(* IEC 61131-3 sources: daoli-st-library/DL_MathData (part 24) *)

(* ---- FC_DL_StatsDevSumSq.st ---- *)
(*
  ============================================================
  组件名 : FC_DL_StatsDevSumSq
  分类   : DL_MathData
  功能   : 定长样本的离差平方和、自由度与方差计算，支持外部给定均值
  开源溯源 : internal-design（本轮无外部代码逐行引用）
             参考语义 : 无外部参考
  复杂度 : C1
  版本   : 1.0.0
  ============================================================
*)

FUNCTION FC_DL_StatsDevSumSq : REAL
VAR_INPUT
    aData        : ARRAY[0..31] OF REAL; // 样本数组，定长三十二 [工程单位] sample array of thirty two fixed slots [engineering unit]
    nCount       : INT; // 有效样本数 1~32 [个] effective sample count from one to thirty two [count]
    rMeanGiven   : REAL; // 外部给定的均值 [工程单位] externally supplied mean [engineering unit]
    bUseGivenMean: BOOL; // 真为使用给定均值，假为按样本自算 use the supplied mean when true
END_VAR
VAR_OUTPUT
    rSs    : REAL; // 离差平方和 [工程单位平方] sum of squared deviations [engineering unit squared]
    rDf    : REAL; // 自由度 [个] degrees of freedom [count]
    rVar   : REAL; // 方差 [工程单位平方] variance [engineering unit squared]
    bValid : BOOL; // 结果有效标志 result validity flag
END_VAR
VAR CONSTANT
    DL_CAP : INT := 32; // 数组容量 [个] array capacity [count]
END_VAR
VAR
    i      : INT := 0; // 遍历游标 [个] walk cursor [count]
    _rMean : REAL := 0.0; // 实际使用的均值 [工程单位] mean actually used [engineering unit]
    _rSum  : REAL := 0.0; // 样本和 [工程单位] sum of the samples [engineering unit]
    _rSs   : REAL := 0.0; // 平方和中间量 [工程单位平方] intermediate sum of squares [engineering unit squared]
    _rDev  : REAL := 0.0; // 单点离差 [工程单位] single deviation [engineering unit]
END_VAR

// 段 1｜出口预置 preset the exit
FC_DL_StatsDevSumSq := 0.0; // 缺省返回零 default zero return
rSs := 0.0; // 平方和预置零 sum of squares preset to zero
rDf := 0.0; // 自由度预置零 freedom preset to zero
rVar := 0.0; // 方差预置零 variance preset to zero
bValid := FALSE; // 计算完成前不认结果 unusable before the calculation
// 段 2｜点数闸与有限闸 count gate and finiteness gate
IF (nCount < 1) OR (nCount > DL_CAP) THEN
    RETURN; // 点数越界即无效 an out of range count is void
END_IF
IF (rMeanGiven <> rMeanGiven) OR ((aData[0] <> aData[0])) THEN
    RETURN; // 均值或首样本非有限即无效 a non finite mean or first sample is void
END_IF
// 段 3｜均值来源选择 the mean source selection
IF bUseGivenMean THEN
    _rMean := rMeanGiven; // 使用外部给定均值 use the supplied mean
ELSE
    _rSum := 0.0; // 样本和清零 clear the sum
    FOR i := 0 TO (nCount - 1) DO
        IF aData[i] <> aData[i] THEN
            RETURN; // 非有限样本拒收 refuse a non finite sample
        END_IF
        _rSum := _rSum + aData[i]; // 样本累加 accumulate the sample
    END_FOR
    _rMean := _rSum / INT_TO_REAL(nCount); // 自算均值，除子为已证正计数 the computed mean over a proven positive count
END_IF
// 段 4｜离差平方和 sum of squared deviations
_rSs := 0.0; // 平方和清零 clear the sum of squares
FOR i := 0 TO (nCount - 1) DO
    IF aData[i] <> aData[i] THEN
        RETURN; // 非有限样本拒收 refuse a non finite sample
    END_IF
    _rDev := aData[i] - _rMean; // 单点离差 single deviation
    _rSs := _rSs + _rDev * _rDev; // 平方累加 accumulate the square
END_FOR
rSs := _rSs; // 平方和落定 land the sum of squares
// 段 5｜自由度与方差自由度闸 freedom and the variance gate
rDf := INT_TO_REAL(nCount - 1); // 自由度取样本数减一 the freedom is the count minus one
IF rDf <= 0.0 THEN
    RETURN; // 自由度非正时方差不可求 a non positive freedom carries no variance
END_IF
rVar := _rSs / rDf; // 方差，除子为已证正自由度 variance over a proven positive freedom
bValid := TRUE; // 结果可用 result usable
FC_DL_StatsDevSumSq := _rSs; // 函数返回离差平方和 return the sum of squares
END_FUNCTION

(* ---- FC_DL_StatsEntropyCalc.st ---- *)
(*==============================================================================
 * 组件名称 : FC_DL_StatsEntropyCalc ｜ 子库 : DL_MathData ｜ v1.0.0 ｜ 2026-11-24
 * 平台     : CODESYS 3.5 / TwinCAT 3 / InoProShop / Machine Expert（纯 IEC，无厂商库）
 * 功能简介 : 香农熵 H = −Σ p·log2(p) [bit]，供直方图分布集中度、缺陷类别混杂度、
 *            多路料仓配比均匀度评估。概率先求和再归一化（q = p / Σp），故入参不要求
 *            严格和为 1（计数直方图可直接喂入）。
 * 契约     : 1 ≤ nCnt ≤ 8、各 p ≥ 0 且有限、Σp > 1.0E-12 → 返回 H ≥ 0、bValid := TRUE；
 *            nCnt 越界、任一 p 为负或非有限、Σp ≤ 1.0E-12（全零/近零，熵无定义）→
 *            返回 0、bError := TRUE、bValid := FALSE。
 * 依赖     : 无 DL_ 内部依赖（R16 自足实现），仅用标准库 LN；log2(p) 以 LN(p)/LN(2) 实现
 * 错误码   : R297 零码位范式：eErr 恒 0，仅以 bError / bValid 表达
 * 红线自检 : R1 零全局 R2 零%I/%Q R3 纯IEC R4 除零前置（Σp 域闸、LN(2) 为常量）+ 跳过 log(0)
 *            R5 双语注释 R6 N/A（无状态机）R7 N/A（无定时器/沿实例）
 *            R10 无类型转换 R11 全声明行分号 R15 标识符零保留字冲突
 *            R17 数组显式定长 ARRAY[1..8]，nCnt 已域闸，无 VLA
 * 遗留假设 : 概率阈值 1.0E-12 以下的项整体跳过（p·log2 p → 0 的极限口径，也避免 LN(0)）；
 *            归一化后才取对数，故入参是计数或百分比皆可；nCnt 之外的数组槽位不参与运算；
 *            H 的量纲为 bit（底数 2），理论上界为 log2(8) = 3.0 bit。
 * 修订历史 : 2026-11-24 R79-B 首版（统计族 2/2）
 *============================================================================*)
FUNCTION FC_DL_StatsEntropyCalc : LREAL
VAR_INPUT
    aProb : ARRAY[1..8] OF LREAL; // 概率或计数数组，元素须 ≥ 0，仅前 nCnt 项参与 [无量纲] / the probability or count vector, only the first nCnt entries are used
    nCnt  : INT := 0;             // 有效元素个数，1..8 [个] / the number of valid entries
END_VAR
VAR_OUTPUT
    eErr   : UDINT; // 错误码，零码位范式恒 0 / error id, always zero under the zero-code rule
    bError : BOOL;  // 个数越界、元素非法或总和近零时为真 / TRUE on a bad count, an illegal entry or a near zero sum
    bValid : BOOL;  // 返回值可用标志 / TRUE when the return value is usable
END_VAR
VAR CONSTANT
    DL_ZERO : LREAL := 0.0;                // 实数零哨兵 [无量纲] / the real zero sentinel
    DL_EPS  : LREAL := 1.0E-12;            // 可忽略概率 / 近零总和阈值 [无量纲] / the negligible probability and near zero sum threshold
    DL_LN2  : LREAL := 0.6931471805599453; // ln2，换底用 [无量纲] / the natural logarithm of two used for the base change
    DL_CNT1 : INT   := 1;                  // 元素个数下界 [个] / the lower entry count bound
    DL_CNT8 : INT   := 8;                  // 元素个数上界 [个] / the upper entry count bound
    DL_ONE  : INT   := 1;                  // 循环起点下标 [无量纲] / the loop start index
    DL_STEP : INT   := 1;                  // 下标步长 [无量纲] / the index step
END_VAR
VAR
    nI    : INT;   // 数组下标 1..nCnt [无量纲] / the array index
    fSum  : LREAL; // 概率总和 Σp [无量纲] / the sum of the probabilities
    fQ    : LREAL; // 归一化概率 p / Σp [无量纲] / the normalised probability
    fH    : LREAL; // 熵累加量 [bit] / the entropy accumulator
END_VAR

// 段 1｜出口预置 / segment 1, preset the exit
FC_DL_StatsEntropyCalc := DL_ZERO;  // 缺省零 / default zero
eErr   := 0;                        // 零码位范式 / zero-code rule
bError := FALSE;                    // 预置无故障 / preset no fault
bValid := FALSE;                    // 域闸前不认返回值 / the return value is unusable until the gates pass

// 段 2｜元素个数域闸：数组定长 1..8，越界下标不可触 / segment 2, the entry count gate
IF (nCnt < DL_CNT1) OR (nCnt > DL_CNT8) THEN
    bError := TRUE;                 // 个数越界 / the count is out of range
    RETURN;                         // 返回 0 / return the preset zero
END_IF

// 段 3｜求和与元素合法性：负概率无意义，非有限入参直接拦 / segment 3, the sum and the entry checks
fSum := DL_ZERO;                    // 总和清零 / clear the sum
FOR nI := DL_ONE TO nCnt DO         // 只遍历有效槽位 / loop over the valid entries only
    IF (aProb[nI] <> aProb[nI]) THEN
        bError := TRUE;             // NaN 元素 / a NaN entry
        RETURN;                     // 返回 0 / return the preset zero
    END_IF
    IF ((aProb[nI] - aProb[nI]) <> DL_ZERO) OR (aProb[nI] < DL_ZERO) THEN
        bError := TRUE;             // Inf 元素或负概率 / an infinite entry or a negative probability
        RETURN;                     // 返回 0 / return the preset zero
    END_IF
    fSum := fSum + aProb[nI];       // 累加 / accumulate
END_FOR

// 段 4｜总和域闸：全零或近零时熵无定义，且归一化会除零 / segment 4, the sum gate
IF fSum <= DL_EPS THEN
    bError := TRUE;                 // 总和近零 / the sum is negligible
    RETURN;                         // 返回 0 / return the preset zero
END_IF
IF (fSum - fSum) <> DL_ZERO THEN    // 溢出成 Inf 的兜底 / the overflow to infinity guard
    bError := TRUE;                 // 总和非有限 / the sum is not finite
    RETURN;                         // 返回 0 / return the preset zero
END_IF

// 段 5｜熵求值：H = −Σ q·log2(q)，q = p / Σp，log2 用 LN(q)/LN(2) / segment 5, the entropy
fH := DL_ZERO;                      // 熵清零 / clear the entropy
FOR nI := DL_ONE TO nCnt DO         // 第二遍：归一化后逐项累加 / second pass over the normalised terms
    IF aProb[nI] > DL_EPS THEN      // 跳过可忽略项，等价 ln(0) 极限且防 log(0) / skip negligible terms to avoid the logarithm of zero
        fQ := aProb[nI] / fSum;     // 归一化（fSum 已证 > 1E-12）/ normalise, the sum is proven positive
        fH := fH - (fQ * (LN(fQ) / DL_LN2));  // 累减 q·log2 q [bit] / subtract the term
    END_IF
END_FOR

// 段 6｜出口 / segment 6, the exit
FC_DL_StatsEntropyCalc := fH;       // 回写熵 [bit] / publish the entropy
bValid := TRUE;                     // 返回值可用 / the return value is usable
END_FUNCTION

(* ---- FC_DL_StatsHistogramBin.st ---- *)
(*==============================================================================
 * 组件名称 : FC_DL_StatsHistogramBin ｜ 子库 : DL_MathData ｜ v1.0.0 ｜ 2026-11-24
 * 平台     : CODESYS 3.5 / TwinCAT 3 / InoProShop / Machine Expert（纯 IEC，无厂商库）
 * 功能简介 : 等宽直方图落桶序号。桶宽 fWidth、桶数 nBins、起点 fMin 给定，
 *            返回 1~nBins 的桶号，供桶计数数组自增（直方图 = 落桶 + 计数两步）。
 *            首尾桶按开区间外延钳位：小于起点归首桶，大于末桶归末桶 ——
 *            线上数据超界不该丢样本，也不该写越界下标。
 * 契约     : 返回 1~nBins；fVal < fMin 返回 1，fVal ≥ 末桶上界返回 nBins；
 *            fWidth ≤ 1.0E-9 或 nBins < 1 返回 0、bError := TRUE（桶结构非法）；
 *            非有限输入返回 0、bError := TRUE。
 * 依赖     : 无 DL_ 内部依赖（R16 自足实现）；Standard.library: TRUNC / ABS
 * 错误码   : R297 零码位范式：eErr 恒 0，仅以 bError / bValid 表达
 * 红线自检 : R1 零全局 R2 零%I/%Q R3 纯IEC R4 桶宽闸防除零、实数上限兜底后才取整防溢出、
 *            NaN 自反判据 ｜ R5 双语注释 R6 N/A（无状态机）R7 N/A（无定时器/沿实例）
 *            R10 标准转换（TRUNC + LREAL_TO_DINT）R11 全声明行分号
 *            R15 标识符零保留字冲突 R18 N/A（无 bReset）
 * 修订历史 : 2026-11-24 R79-A 首版（统计扩展族 7/8）
 *============================================================================*)
FUNCTION FC_DL_StatsHistogramBin : DINT
VAR_INPUT
    fVal    : LREAL;    // 待落桶样本 [工程单位] / sample to place into a bin [engineering unit]
    fMin    : LREAL;    // 首桶下界（含） [工程单位] / lower edge of the first bin, inclusive [engineering unit]
    fWidth  : LREAL;    // 桶宽，须 > 0 [工程单位] / bin width, must be positive [engineering unit]
    nBins   : INT;      // 桶数，须 ≥ 1 [个] / bin count, at least one [count]
END_VAR
VAR_OUTPUT
    eErr    : UDINT;    // 错误码，零码位范式恒 0 / error id, always zero under the zero-code rule
    bError  : BOOL;     // 桶结构非法或输入非有限为真 / TRUE on an illegal bin structure or non finite inputs
    bValid  : BOOL;     // 结果可用标志 / result usable flag
END_VAR
VAR CONSTANT
    DL_WIDTH_MIN : LREAL := 1.0E-9;     // 桶宽下限，低于它判结构非法 [工程单位] / width floor below which the structure is illegal
    DL_FIN_LIM   : LREAL := 1.0E308;    // 有限性上界 [工程单位] / finiteness ceiling
    DL_ONE       : DINT := 1;           // 首桶号与下标偏移 [个] / the first bin number [count]
    DL_ZERO      : DINT := 0;           // 整数零哨兵，代表非法 / integer zero sentinel meaning illegal
    DL_ZERO_L    : LREAL := 0.0;        // 实数零哨兵 / real zero sentinel
END_VAR
VAR
    fOffset : LREAL;    // 样本相对首桶下界的偏移 [工程单位] / offset of the sample from the first lower edge
    fIdx    : LREAL;    // 零基桶序号实数形式 [个] / zero based bin index as a real number
    nBin    : DINT;     // 一基桶序号 [个] / one based bin number [count]
END_VAR

// 段 1｜出口预置：0 为非法桶号 / segment 1, preset the exit with the illegal bin number
FC_DL_StatsHistogramBin := DL_ZERO;     // 缺省非法 / default illegal
eErr   := 0;                            // 零码位范式 / zero-code rule
bError := FALSE;                        // 预置无故障 / preset no fault
bValid := FALSE;                        // 域闸前不认结果 / unusable until the gates pass

// 段 2｜桶结构闸与输入闸：桶宽、桶数、三个实数的有限性 / segment 2, the structure and finiteness gates
IF nBins < DL_ONE THEN
    bError := TRUE;                     // 桶数非法 / the bin count is illegal
    RETURN;
END_IF
IF fWidth < DL_WIDTH_MIN THEN
    bError := TRUE;                     // 桶宽非正或近零，落桶除零不可达 / the width is not positive, division is blocked here
    RETURN;
END_IF
IF (fVal <> fVal) OR (fMin <> fMin) OR (fWidth <> fWidth) THEN
    bError := TRUE;                     // 含非数输入 / a not a number input was seen
    RETURN;
END_IF
IF (ABS(fVal) > DL_FIN_LIM) OR (ABS(fMin) > DL_FIN_LIM) THEN
    bError := TRUE;                     // 量级非有限 / a magnitude is not finite
    RETURN;
END_IF

// 段 3｜偏移与首桶钳位：低于起点一律归首桶 / segment 3, the offset and the first bin clamp
fOffset := fVal - fMin;                 // 相对偏移 / the relative offset
IF fOffset < DL_ZERO_L THEN
    FC_DL_StatsHistogramBin := DL_ONE;  // 首桶钳位 / clamp into the first bin
    bValid := TRUE;
    RETURN;
END_IF

// 段 4｜零基序号：先做实数上限兜底再取整，防取整溢出 / segment 4, the real bound before the truncation
fIdx := fOffset / fWidth;               // 分母已证 ≥ 容差 / the divisor is proven to be at least the floor
IF fIdx >= INT_TO_LREAL(nBins) THEN
    FC_DL_StatsHistogramBin := INT_TO_DINT(nBins);      // 末桶钳位，越界样本不丢 / clamp into the last bin
    bValid := TRUE;
    RETURN;
END_IF
nBin := LREAL_TO_DINT(TRUNC(fIdx)) + DL_ONE;            // 零基转一基 / zero based to one based

// 段 5｜出口：档位已证落在 1..nBins / segment 5, the bin is proven to be inside the range
FC_DL_StatsHistogramBin := nBin;        // 桶号 / the bin number
bValid := TRUE;                         // 结果可用 / the result is usable
END_FUNCTION

(* ---- FC_DL_StatsPercentileRankFixed.st ---- *)
(*==============================================================================
 * 组件名称 : FC_DL_StatsPercentileRankFixed ｜ 子库 : DL_MathData ｜ v1.0.0 ｜ 2026-11-24
 * 平台     : CODESYS 3.5 / TwinCAT 3 / InoProShop / Machine Expert（纯 IEC，无厂商库）
 * 功能简介 : 定长样本的分位数（最近秩法 nearest-rank）—— 先升序排序，
 *            rank = ceil(pct/100 × n) 并钳到 [1, n]，返回第 rank 个样本。
 *            最近秩法不插值，返回的一定是真实测得的样本值，HMI 展示与判定门槛
 *            不会因插值出现「从未测到的数」。用于节拍 P95、温度 P99 等分位统计。
 * 契约     : 返回分位数（必为样本之一）；nCnt < 1 时返回 0 且 bError := TRUE；
 *            nCnt > 10 钳到 10；fPct 越界钳到 [0,100]（钳位不报错，属正常输入整形）。
 *            排序用自实现插入排序，数组定长 ARRAY[1..10]（R17）。
 * 依赖     : 无 DL_ 内部依赖（R16 自足实现）；Standard.library: CEIL
 * 错误码   : R297 零码位范式：eErr 恒 0，仅以 bError / bValid 表达
 * 红线自检 : R1 零全局 R2 零%I/%Q R3 纯IEC R4 点数与百分位双钳位、秩再钳到 [1,n]，
 *            下标恒合法 ｜ R5 双语注释 R6 N/A（无状态机）R7 N/A（无定时器/沿实例）
 *            R10 标准转换 R11 全声明行分号 R15 标识符零保留字冲突
 *            R17 定长数组 R18 N/A（无 bReset）
 * 遗留假设 : 最近秩法在 pct = 0 时 rank = 0 会钳到 1（返回最小值），与教科书「P0」口径一致。
 * 修订历史 : 2026-11-24 R79-A 首版（统计扩展族 5/8）
 *============================================================================*)
FUNCTION FC_DL_StatsPercentileRankFixed : LREAL
VAR_INPUT
    aVals   : ARRAY[1..10] OF LREAL;    // 样本数组，1..10 定长 [工程单位] / sample array of fixed length [engineering unit]
    nCnt    : INT;                      // 有效样本数，1~10，越界钳位 [个] / effective sample count from one to ten, clamped [count]
    fPct    : LREAL;                    // 百分位 0~100，越界钳位 [%] / percentile from zero to one hundred, clamped [%]
END_VAR
VAR_OUTPUT
    eErr    : UDINT;                    // 错误码，零码位范式恒 0 / error id, always zero under the zero-code rule
    bError  : BOOL;                     // 有效样本数为零为真 / TRUE when no usable sample exists
    bValid  : BOOL;                     // 结果可用标志 / result usable flag
END_VAR
VAR CONSTANT
    DL_PTS_MAX : INT := 10;             // 样本定长上限 [个] / fixed sample capacity [count]
    DL_PTS_MIN : INT := 1;              // 最少样本数 [个] / minimum sample count [count]
    DL_ONE     : INT := 1;              // 数组首下标与秩下界 [个] / first index and the lower rank bound [count]
    DL_TWO     : INT := 2;              // 插入排序的起始下标 [个] / starting index of the insertion sort [count]
    DL_PCT_MIN : LREAL := 0.0;          // 百分位下界 [%] / lower percentile bound [%]
    DL_PCT_MAX : LREAL := 100.0;        // 百分位上界 [%] / upper percentile bound [%]
    DL_PCT_DIV : LREAL := 100.0;        // 百分制换算除数 [%] / percentile scale divisor [%]
    DL_ZERO_L  : LREAL := 0.0;          // 实数零哨兵 [工程单位] / real zero sentinel [engineering unit]
END_VAR
VAR
    aBuf    : ARRAY[1..10] OF LREAL;    // 排序后的样本副本 [工程单位] / sorted copy of the samples [engineering unit]
    nUse    : INT;                      // 钳位后的有效点数 [个] / effective point count after clamping [count]
    nRank   : INT;                      // 最近秩 1~nUse [个] / the nearest rank from one to the count [count]
    i       : INT;                      // 外层游标 [个] / outer cursor [count]
    j       : INT;                      // 内层游标 [个] / inner cursor [count]
    fKey    : LREAL;                    // 插入排序待插值 [工程单位] / key of the insertion sort [engineering unit]
    fPctUse : LREAL;                    // 钳位后的百分位 [%] / effective percentile after clamping [%]
    fRank   : LREAL;                    // 秩的实数中间量 [个] / the rank as a real number [count]
END_VAR

// 段 1｜出口预置 / segment 1, preset the exit
FC_DL_StatsPercentileRankFixed := DL_ZERO_L;    // 缺省 0 / default zero
eErr    := 0;                                   // 零码位范式 / zero-code rule
bError  := FALSE;                               // 预置无故障 / preset no fault
bValid  := FALSE;                               // 计算完成前不认结果 / unusable until the rank walk ends

// 段 2｜点数钳位与百分位整形 / segment 2, clamp the count and normalise the percentile
nUse := nCnt;
IF nUse > DL_PTS_MAX THEN
    nUse := DL_PTS_MAX;
END_IF
IF nUse < DL_PTS_MIN THEN
    bError := TRUE;                             // 无样本可统计 / no sample to scan
    RETURN;
END_IF
fPctUse := fPct;
IF (fPctUse <> fPctUse) OR (fPctUse < DL_PCT_MIN) THEN
    fPctUse := DL_PCT_MIN;                      // 非数或过小按 0 处理 / a not a number or an undershoot becomes zero
ELSIF fPctUse > DL_PCT_MAX THEN
    fPctUse := DL_PCT_MAX;                      // 过大按 100 处理 / an overshoot becomes one hundred
END_IF

// 段 3｜拷贝并插入排序：升序，秩直接映射到下标 / segment 3, copy and insertion sort
FOR i := DL_ONE TO nUse DO
    aBuf[i] := aVals[i];                        // 拷贝，保持入参只读 / copy so the input stays read only
END_FOR
FOR i := DL_TWO TO nUse DO
    fKey := aBuf[i];
    j    := i - DL_ONE;
    WHILE (j >= DL_ONE) AND (aBuf[j] > fKey) DO
        aBuf[j + DL_ONE] := aBuf[j];            // 后移空位 / shift right to open a slot
        j := j - DL_ONE;
    END_WHILE
    aBuf[j + DL_ONE] := fKey;                   // 落位 / drop the key in place
END_FOR

// 段 4｜最近秩：ceil(pct/100 × n)，再钳到 [1, n] / segment 4, the nearest rank
fRank := CEIL((fPctUse / DL_PCT_DIV) * INT_TO_LREAL(nUse));    // 向上取整，整数域内无插值误差 / round up, no interpolation error
nRank := LREAL_TO_DINT(fRank);                                 // 转整数秩 / convert to an integer rank
IF nRank < DL_ONE THEN
    nRank := DL_ONE;                                           // 秩下界钳位 / clamp the lower rank bound
ELSIF nRank > nUse THEN
    nRank := nUse;                                             // 秩上界钳位 / clamp the upper rank bound
END_IF

// 段 5｜出口：秩已证落在 [1, nUse]，下标安全 / segment 5, the rank is proven legal
FC_DL_StatsPercentileRankFixed := aBuf[nRank];      // 该分位的实测样本值 / the measured sample at that percentile
bValid := TRUE;                                     // 结果可用 / the result is usable
END_FUNCTION

(* ---- FC_DL_StatsPooledStd.st ---- *)
(*
  ============================================================
  组件名 : FC_DL_StatsPooledStd
  分类   : DL_MathData
  功能   : 两组样本的合并方差与合并标准差计算，按自由度加权
  开源溯源 : internal-design（本轮无外部代码逐行引用）
             参考语义 : 无外部参考
  复杂度 : C1
  版本   : 1.0.0
  ============================================================
*)

FUNCTION FC_DL_StatsPooledStd : REAL
VAR_INPUT
    rVar1 : REAL; // 第一组样本方差 [工程单位平方] variance of the first group [engineering unit squared]
    rVar2 : REAL; // 第二组样本方差 [工程单位平方] variance of the second group [engineering unit squared]
    n1    : INT; // 第一组样本数 [个] first group sample count [count]
    n2    : INT; // 第二组样本数 [个] second group sample count [count]
END_VAR
VAR_OUTPUT
    rPooledVar : REAL; // 合并方差 [工程单位平方] pooled variance [engineering unit squared]
    rPooledStd : REAL; // 合并标准差 [工程单位] pooled standard deviation [engineering unit]
    nDf        : INT; // 合并自由度 [个] pooled degrees of freedom [count]
    bValid     : BOOL; // 结果有效标志 result validity flag
END_VAR
VAR
    _bFin : BOOL := FALSE; // 两实数输入有限性判定 finiteness verdict of both real inputs
    _rNum : REAL := 0.0; // 自由度加权分子 [工程单位平方] weighted numerator [engineering unit squared]
    _rVar : REAL := 0.0; // 合并方差中间量 [工程单位平方] intermediate pooled variance [engineering unit squared]
    _rStd : REAL := 0.0; // 合并标准差中间量 [工程单位] intermediate pooled deviation [engineering unit]
END_VAR

// 段 1｜出口预置 preset the exit
FC_DL_StatsPooledStd := 0.0; // 缺省返回零 default zero return
rPooledVar := 0.0; // 合并方差预置零 pooled variance preset to zero
rPooledStd := 0.0; // 合并标准差预置零 pooled deviation preset to zero
nDf := 0; // 自由度预置零 degrees of freedom preset to zero
bValid := FALSE; // 计算完成前不认结果 unusable before the calculation
// 段 2｜非有限闸 finiteness gate
_bFin := (rVar1 = rVar1) AND (rVar2 = rVar2); // 两输入自反判定 self comparison of both inputs
IF NOT _bFin THEN
    RETURN; // 非有限即无效 non finite means invalid
END_IF
// 段 3｜方差方向闸与样本数闸 variance direction gate and count gate
IF (rVar1 < 0.0) OR (rVar2 < 0.0) THEN
    RETURN; // 负方差属计算异常 a negative variance is an illegal input
END_IF
IF (n1 < 1) OR (n2 < 1) THEN
    RETURN; // 组样本数非正无法加权 a non positive group count cannot be weighted
END_IF
// 段 4｜自由度与合并方差 degrees of freedom and the pooled variance
nDf := n1 + n2 - 2; // 合并自由度 pooled degrees of freedom
IF nDf <= 0 THEN
    RETURN; // 自由度非正无法求方差 a non positive freedom cannot carry a variance
END_IF
_rNum := INT_TO_REAL(n1 - 1) * rVar1 + INT_TO_REAL(n2 - 1) * rVar2; // 自由度加权分子 weighted numerator
_rVar := _rNum / INT_TO_REAL(nDf); // 合并方差，除子已证为正 pooled variance over a proven positive divisor
rPooledVar := _rVar; // 合并方差落定 land the pooled variance
// 段 5｜合并标准差与出口 pooled deviation and the exit
_rStd := SQRT(_rVar); // 方差开方得标准差 the square root of the variance
rPooledStd := _rStd; // 合并标准差落定 land the pooled deviation
bValid := TRUE; // 结果可用 result usable
FC_DL_StatsPooledStd := _rStd; // 函数返回合并标准差 return the pooled deviation
END_FUNCTION

(* ---- FC_DL_StatsRangeCalc.st ---- *)
(*
  ============================================================
  组件名 : FC_DL_StatsRangeCalc
  分类   : DL_MathData
  功能   : 定长样本的极差统计，返回最小值、最大值与极差
  开源溯源 : internal-design（本轮无外部代码逐行引用）
             参考语义 : 无外部参考
  复杂度 : C1
  版本   : 1.0.0
  ============================================================
*)

FUNCTION FC_DL_StatsRangeCalc : REAL
VAR_INPUT
    aData  : ARRAY[0..31] OF REAL; // 样本数组，定长三十二 [工程单位] sample array of thirty two fixed slots [engineering unit]
    nCount : INT; // 有效样本数 1~32 [个] effective sample count from one to thirty two [count]
END_VAR
VAR_OUTPUT
    rRange : REAL; // 极差 [工程单位] range [engineering unit]
    rMin   : REAL; // 最小值 [工程单位] minimum [engineering unit]
    rMax   : REAL; // 最大值 [工程单位] maximum [engineering unit]
    nUsed  : INT; // 实际参与统计的点数 [个] point count actually used [count]
    bValid : BOOL; // 结果有效标志 result validity flag
END_VAR
VAR CONSTANT
    DL_CAP  : INT := 32; // 数组容量 [个] array capacity [count]
END_VAR
VAR
    i     : INT := 0; // 遍历游标 [个] walk cursor [count]
    _rMin : REAL := 0.0; // 最小值中间量 [工程单位] intermediate minimum [engineering unit]
    _rMax : REAL := 0.0; // 最大值中间量 [工程单位] intermediate maximum [engineering unit]
    _bFin : BOOL := FALSE; // 当前样本有限性判定 finiteness verdict of the current sample
END_VAR

// 段 1｜出口预置 preset the exit
FC_DL_StatsRangeCalc := 0.0; // 缺省返回零 default zero return
rRange := 0.0; // 极差预置零 range preset to zero
rMin := 0.0; // 最小值预置零 minimum preset to zero
rMax := 0.0; // 最大值预置零 maximum preset to zero
nUsed := 0; // 参与点数预置零 used count preset to zero
bValid := FALSE; // 计算完成前不认结果 unusable before the calculation
// 段 2｜点数闸 sample count gate
IF (nCount < 1) OR (nCount > DL_CAP) THEN
    RETURN; // 点数越界即无效 an out of range count is void
END_IF
// 段 3｜初值取首样本 the first sample seeds both bounds
_bFin := (aData[0] = aData[0]); // 首样本自反判定 self comparison of the first sample
IF NOT _bFin THEN
    RETURN; // 首样本非有限即无效 a non finite seed is void
END_IF
_rMin := aData[0]; // 最小值初值取首样本 the minimum starts at the first sample
_rMax := aData[0]; // 最大值初值取首样本 the maximum starts at the first sample
// 段 4｜单趟遍历求双向极值 single pass over both bounds
FOR i := 1 TO (nCount - 1) DO
    IF aData[i] <> aData[i] THEN
        RETURN; // 非有限样本拒收，出口回零点 refuse a non finite sample and return the zero outlet
    END_IF
    IF aData[i] < _rMin THEN
        _rMin := aData[i]; // 刷新最小值 refresh the minimum
    END_IF
    IF aData[i] > _rMax THEN
        _rMax := aData[i]; // 刷新最大值 refresh the maximum
    END_IF
END_FOR
// 段 5｜极差与出口 range and the exit
rMin := _rMin; // 最小值落定 land the minimum
rMax := _rMax; // 最大值落定 land the maximum
rRange := _rMax - _rMin; // 极差为最大值减最小值 the range is the maximum minus the minimum
nUsed := nCount; // 参与点数落定 land the used count
bValid := TRUE; // 结果可用 result usable
FC_DL_StatsRangeCalc := rRange; // 函数返回极差 return the range
END_FUNCTION

(* ---- FC_DL_StatsRunLengthMax.st ---- *)
(*==============================================================================
 * 组件名称 : FC_DL_StatsRunLengthMax ｜ 子库 : DL_MathData ｜ v1.0.0 ｜ 2026-11-24
 * 平台     : CODESYS 3.5 / TwinCAT 3 / InoProShop / Machine Expert（纯 IEC，无厂商库）
 * 功能简介 : 定长样本的最长「连续同值游程」（run length）长度。相邻两样本差值
 *            不超过 fTol 即视为同值，游程在容差内延续。用于：称重稳定判定、
 *            光电信号连续遮挡时长、清洗液浓度平台段长度、批次工艺稳态持续时间。
 * 契约     : 返回最长游程长度（1~nCnt）；nCnt < 1 时返回 0 且 bError := TRUE；
 *            nCnt > 10 钳到 10；fTol 取绝对值（负容差按同值正容差处理），
 *            非有限 fTol 返回 0 且 bError := TRUE。数组定长 ARRAY[1..10]（R17）。
 * 依赖     : 无 DL_ 内部依赖（R16 自足实现）；Standard.library: ABS
 * 错误码   : R297 零码位范式：eErr 恒 0，仅以 bError / bValid 表达
 * 红线自检 : R1 零全局 R2 零%I/%Q R3 纯IEC R4 点数先钳位后扫描、容差常量化、
 *            浮点差值比较走 ABS 容差不用等号、NaN 自反判据 ｜ R5 双语注释
 *            R6 N/A（无状态机）R7 N/A（无定时器/沿实例）R10 无类型转换
 *            R11 全声明行分号 R15 标识符零保留字冲突 R17 定长数组 R18 N/A（无 bReset）
 * 修订历史 : 2026-11-24 R79-A 首版（统计扩展族 8/8）
 *============================================================================*)
FUNCTION FC_DL_StatsRunLengthMax : DINT
VAR_INPUT
    aVals   : ARRAY[1..10] OF LREAL;    // 样本数组，1..10 定长 [工程单位] / sample array of fixed length [engineering unit]
    nCnt    : INT;                      // 有效样本数，1~10，越界钳位 [个] / effective sample count from one to ten, clamped [count]
    fTol    : LREAL;                    // 同值容差，取绝对值使用 [工程单位] / equality tolerance, used as a magnitude [engineering unit]
END_VAR
VAR_OUTPUT
    eErr    : UDINT;                    // 错误码，零码位范式恒 0 / error id, always zero under the zero-code rule
    bError  : BOOL;                     // 无样本或容差非有限为真 / TRUE when no sample exists or the tolerance is not finite
    bValid  : BOOL;                     // 结果可用标志 / result usable flag
END_VAR
VAR CONSTANT
    DL_PTS_MAX : INT := 10;             // 样本定长上限 [个] / fixed sample capacity [count]
    DL_PTS_MIN : INT := 1;              // 最少样本数 [个] / minimum sample count [count]
    DL_ONE     : INT := 1;              // 数组首下标与最短游程 [个] / first index and the shortest possible run [count]
    DL_ZERO    : INT := 0;              // 整数零哨兵 / integer zero sentinel
    DL_FIN_LIM : LREAL := 1.0E308;      // 有限性上界 [工程单位] / finiteness ceiling [engineering unit]
END_VAR
VAR
    nUse    : INT;                      // 钳位后的有效点数 [个] / effective point count after clamping [count]
    nRun    : INT;                      // 当前游程长度 [个] / the run being measured [count]
    nBest   : INT;                      // 历史最长游程 [个] / the longest run seen so far [count]
    i       : INT;                      // 遍历游标，从第 2 点起 [个] / loop cursor starting at the second point [count]
    fTolUse : LREAL;                    // 生效容差 [工程单位] / effective tolerance [engineering unit]
    fDiff   : LREAL;                    // 相邻样本差值 [工程单位] / difference of neighbouring samples [engineering unit]
END_VAR

// 段 1｜出口预置 / segment 1, preset the exit
FC_DL_StatsRunLengthMax := DL_ZERO;     // 缺省 0 / default zero
eErr   := 0;                            // 零码位范式 / zero-code rule
bError := FALSE;                        // 预置无故障 / preset no fault
bValid := FALSE;                        // 计算完成前不认结果 / unusable until the scan ends

// 段 2｜点数钳位与容差整形 / segment 2, clamp the count and normalise the tolerance
nUse := nCnt;
IF nUse > DL_PTS_MAX THEN
    nUse := DL_PTS_MAX;                 // 钳到定长上限 / clamp to the fixed capacity
END_IF
IF nUse < DL_PTS_MIN THEN
    bError := TRUE;                     // 无样本可扫描 / no sample to scan
    RETURN;
END_IF
IF (fTol <> fTol) OR (ABS(fTol) > DL_FIN_LIM) THEN
    bError := TRUE;                     // 容差非数或无穷 / the tolerance is not finite
    RETURN;
END_IF
fTolUse := ABS(fTol);                   // 负容差按同值正容差处理 / a negative tolerance folds to its magnitude

// 段 3｜首点起算：单个样本本身构成游程 1 / segment 3, the first sample seeds a run of one
nRun  := DL_ONE;
nBest := DL_ONE;

// 段 4｜单趟扫描：差值在容差内则游程加一，否则重新起算 / segment 4, one pass over the neighbours
FOR i := (DL_ONE + DL_ONE) TO nUse DO
    fDiff := ABS(aVals[i] - aVals[i - DL_ONE]);     // 相邻差值 / neighbouring difference
    IF fDiff <= fTolUse THEN
        nRun := nRun + DL_ONE;                      // 游程延续 / the run continues
        IF nRun > nBest THEN
            nBest := nRun;                          // 刷新最长 / refresh the record
        END_IF
    ELSE
        nRun := DL_ONE;                             // 新值起算新游程 / a new value starts a new run
    END_IF
END_FOR

// 段 5｜出口：nBest 已证落在 1..nUse / segment 5, the record is proven to be inside the range
FC_DL_StatsRunLengthMax := nBest;       // 最长游程 / the longest run
bValid := TRUE;                         // 结果可用 / the result is usable
END_FUNCTION

(* ---- FC_DL_StatsZScoreClamp.st ---- *)
(*==============================================================================
 * 组件名称 : FC_DL_StatsZScoreClamp ｜ 子库 : DL_MathData ｜ v1.0.0 ｜ 2026-11-24
 * 平台     : CODESYS 3.5 / TwinCAT 3 / InoProShop / Machine Expert（纯 IEC，无厂商库）
 * 功能简介 : 标准化偏差（z 分数）计算并对称限幅。z = (x − mean) / std，再钳到 ±fClamp。
 *            限幅的意义：异常样本的 z 可能上千，直接送 PID 或神经网络会把输出顶到饱和；
 *            钳到 ±3~±5 既保留「异常」信息又不炸控制器。
 * 契约     : 返回 z（已钳位）；fStd < 1.0E-9 时返回 0（除零结构性不可达，零标准差无 z 可言）；
 *            fClamp ≤ 0 时按 1.0 处理（限幅必须为正，否则钳位区间退化为一点）；
 *            任一输入为 NaN 或非有限值时返回 0、bError := TRUE、bValid := FALSE。
 * 依赖     : 无 DL_ 内部依赖（R16 自足实现）；Standard.library: ABS
 * 错误码   : R297 零码位范式：eErr 恒 0，仅以 bError / bValid 表达
 * 红线自检 : R1 零全局 R2 零%I/%Q R3 纯IEC R4 除零前置（std 阈值闸）、NaN 自反判据、
 *            无穷上界、fClamp 非正回退 ｜ R5 双语注释 R6 N/A（无状态机）
 *            R7 N/A（无定时器/沿实例）R10 无类型转换 R11 全声明行分号
 *            R15 标识符零保留字冲突 R18 N/A（无 bReset）
 * 修订历史 : 2026-11-24 R79-A 首版（统计扩展族 6/8）
 *============================================================================*)
FUNCTION FC_DL_StatsZScoreClamp : LREAL
VAR_INPUT
    fVal     : LREAL;   // 待标准化样本 [工程单位] / sample to standardise [engineering unit]
    fMean    : LREAL;   // 总体均值 [工程单位] / population mean [engineering unit]
    fStd     : LREAL;   // 总体标准差 [工程单位] / population standard deviation [engineering unit]
    fClamp   : LREAL;   // 对称限幅幅值，须 > 0，非正按 1.0 [无量纲] / symmetric clamp magnitude, non positive falls back to one
END_VAR
VAR_OUTPUT
    eErr     : UDINT;   // 错误码，零码位范式恒 0 / error id, always zero under the zero-code rule
    bError   : BOOL;    // 输入含非有限值为真 / TRUE when an input is not finite
    bValid   : BOOL;    // 结果可用标志 / result usable flag
    bClamped : BOOL;    // 本次结果被限幅为真 / TRUE when the result hit the clamp
END_VAR
VAR CONSTANT
    DL_EPS      : LREAL := 1.0E-9;      // 标准差下限，低于它按零标准差处理 [工程单位] / deviation floor below which the spread counts as zero
    DL_FIN_LIM  : LREAL := 1.0E308;     // 有限性上界 [工程单位] / finiteness ceiling
    DL_CLAMP_DEF : LREAL := 1.0;        // 限幅回退值，非正输入时使用 [无量纲] / clamp fallback used for non positive inputs
    DL_ZERO_L   : LREAL := 0.0;         // 实数零哨兵 / real zero sentinel
END_VAR
VAR
    fClampUse : LREAL;  // 生效限幅幅值，恒为正 [无量纲] / effective clamp magnitude, always positive
    fZ        : LREAL;  // 未限幅的 z 分数 [无量纲] / the raw z score
END_VAR

// 段 1｜出口预置 / segment 1, preset the exit
FC_DL_StatsZScoreClamp := DL_ZERO_L;    // 缺省 z=0 / default z of zero
eErr     := 0;                          // 零码位范式 / zero-code rule
bError   := FALSE;                      // 预置无故障 / preset no fault
bValid   := FALSE;                      // 计算完成前不认结果 / unusable until the computation ends
bClamped := FALSE;                      // 预置未限幅 / preset unclamped

// 段 2｜非有限闸：四个入参逐一验 NaN 与量级 / segment 2, the non finite gate
IF (fVal <> fVal) OR (fMean <> fMean) OR (fStd <> fStd) OR (fClamp <> fClamp) THEN
    bError := TRUE;                     // 含非数输入 / a not a number input was seen
    RETURN;
END_IF
IF (ABS(fVal) > DL_FIN_LIM) OR (ABS(fMean) > DL_FIN_LIM) OR (ABS(fStd) > DL_FIN_LIM) OR (ABS(fClamp) > DL_FIN_LIM) THEN
    bError := TRUE;                     // 量级非有限 / a magnitude is not finite
    RETURN;
END_IF

// 段 3｜限幅幅值整形：非正按 1.0，取绝对值后恒正 / segment 3, normalise the clamp magnitude
fClampUse := ABS(fClamp);
IF fClampUse < DL_EPS THEN
    fClampUse := DL_CLAMP_DEF;          // 退化限幅回退 1.0 / a degenerate clamp falls back to one
END_IF

// 段 4｜零标准差闸：结构性除零在此拦下 / segment 4, the zero deviation gate
IF fStd < DL_EPS THEN
    bValid := TRUE;                     // z 定义为 0，结论可用 / a zero spread yields z of zero, a usable verdict
    RETURN;                             // 返回 0 / return zero
END_IF

// 段 5｜z 分数与对称限幅：分母已证 ≥ 容差 / segment 5, the z score and the symmetric clamp
fZ := (fVal - fMean) / fStd;            // 标准化偏差 / the standardised deviation
IF fZ > fClampUse THEN
    fZ       := fClampUse;              // 上限幅 / clamp on the upper side
    bClamped := TRUE;
ELSIF fZ < -fClampUse THEN
    fZ       := -fClampUse;             // 下限幅 / clamp on the lower side
    bClamped := TRUE;
END_IF

// 段 6｜出口 / segment 6, exit
FC_DL_StatsZScoreClamp := fZ;           // 限幅后的 z / the clamped z score
bValid := TRUE;                         // 结果可用 / the result is usable
END_FUNCTION

(* ---- FC_DL_StringConcatEx.st ---- *)
(*
    FC_DL_StringConcatEx —— 安全拼接防御包装（超 255 截断显式置 bTruncated，R37 范式）
    ------------------------------------------------------------------
    分类      : DL_MathData / String
    前缀      : FC_DL_
    版本      : 1.0.0
    溯源      : IEC 61131-3 标准语义的道莅防御性实现
                （内部委托平台内建函数，外围统一错误码/钳位/双语文档；
                  未复制任何闭源厂商源码，参考实现仅限 MIT/Apache 许可）
    平台      : 纯 IEC 61131-3，CODESYS / TwinCAT / InoProShop 通用
    作者      : 道莅代码库 · PLC编程专家（R15）
    ------------------------------------------------------------------
    功能说明  : 将 sA 与 sB 拼接到 sResult。严禁直接 CONCAT 后不判长的
                静默截断：先锁存两串有效长度，总长 > 255 时按 R37 范式
                先置 VAR_OUTPUT bTruncated=TRUE 与 eErr=16#0001_0277 再钳位
                （B 段配额 = 255 - A 段长），杜绝静默回夹。复制采用逐字
                符 FOR 循环（跨平台口径），每轮带 255 越界 EXIT 守卫，
                复制后显式写空字符终止符。返回值 TRUE 表示已执行完成。
    错误码    : 0000 正常 / 16#0001_0277 上溢下溢（总长超 255，已显式截断，bTruncated=TRUE）
    修订记录  : 2026-11-16 v1.0.0 首次入库（R15）
*)
FUNCTION FC_DL_StringConcatEx : BOOL
VAR_INPUT
    sA : STRING(255); // 拼接前段 [字符] / front part of the concatenation [chars]
    sB : STRING(255); // 拼接后段 [字符] / rear part of the concatenation [chars]
END_VAR
VAR_OUTPUT
    sResult    : STRING(255); // 结果串 [字符]，A 段接 B 段 / result string [chars], front part followed by rear part
    eErr : UDINT; // 错误码，0=正常，2=超 255 显式截断 / error id, 0=ok, 2=explicit truncation at the 255 cap
    bError     : BOOL; // 是否出错，eErr 非 0 时为 TRUE / error flag, TRUE when eErr is nonzero
    bValid     : BOOL; // 输出是否有效可用，截断降级时为 FALSE / output valid, FALSE for truncated degraded results
    bTruncated : BOOL; // 截断标志，发生 255 截断时 TRUE（R37 范式） / truncation flag, TRUE when the 255 cap truncated content, R37 paradigm
END_VAR
VAR
    nI     : INT; // 循环索引 [字符位序]，1 基 / loop index [char position], 1-based
    nLenA  : INT; // 锁存的 A 段有效长度 [字符] / latched effective length of the front part [chars]
    nLenB  : INT; // 锁存的 B 段有效长度 [字符] / latched effective length of the rear part [chars]
    nTotal : INT; // 拼接总长 [字符] / total concatenated length [chars]
    nUseB  : INT; // B 段实际复制数 [字符]，受 255 配额钳制 / chars actually copied from the rear part [chars], clamped by the 255 quota
END_VAR
VAR CONSTANT
    DL_CC_MAX : INT := 255; // 串型上限 [字符] / string type cap [chars]
END_VAR

// 段 1｜返回值与输出预置，任何早退路径不留脏码 / segment 1, preset return value and outputs
FC_DL_StringConcatEx := TRUE; // 返回值预置 TRUE（已执行口径） / preset return to TRUE, executed semantics
sResult              := ''; // 结果串预置空串 / preset result to the empty string
eErr             := 16#0000_0000; // 错误码预置正常 / preset error id to ok
bError               := FALSE; // 错误标志预置无错 / preset error flag to FALSE
bValid               := TRUE; // 有效标志预置可用 / preset valid flag to TRUE
bTruncated           := FALSE; // 截断标志预置无截断 / preset truncation flag to FALSE

// 段 2｜两段有效长度各一次锁存（空字符截止扫描 + 255 越界守卫） / segment 2, latch both effective lengths once
nI    := 1; // 索引起始 [字符位序] / index start
nLenA := 0; // A 段长度预置 [字符] / preset front length
WHILE nI <= DL_CC_MAX DO
    IF nI > DL_CC_MAX THEN   (* 越界守卫（双重保险） EN: overrun guard *)
        EXIT;
    END_IF
    IF sA[nI] = '$00' THEN   (* A 段首个空字符即串结束 EN: first null char ends the front part *)
        EXIT;
    END_IF
    nLenA := nI; // 记录 A 段最后非空位序 [字符] / record the last non-null position
    nI    := nI + 1; // 每轮自增 / per-iteration increment
END_WHILE
nI    := 1; // 索引复位 / reset index
nLenB := 0; // B 段长度预置 [字符] / preset rear length
WHILE nI <= DL_CC_MAX DO
    IF nI > DL_CC_MAX THEN   (* 越界守卫（双重保险） EN: overrun guard *)
        EXIT;
    END_IF
    IF sB[nI] = '$00' THEN   (* B 段首个空字符即串结束 EN: first null char ends the rear part *)
        EXIT;
    END_IF
    nLenB := nI; // 记录 B 段最后非空位序 [字符] / record the last non-null position
    nI    := nI + 1; // 每轮自增 / per-iteration increment
END_WHILE

// 段 3｜255 截断闸（R37 范式：先判定后写入，严禁静默回夹） / segment 3, the 255 truncation gate, R37 paradigm, decide before writing, silent clipping forbidden
nTotal := nLenA + nLenB; // 拼接总长 [字符] / total length
IF nTotal > DL_CC_MAX THEN
    nUseB := DL_CC_MAX - nLenA; // B 段配额 = 255 减 A 段长，可为 0 / rear quota = 255 minus front length, may be zero
    bTruncated := TRUE; // 显式置截断标志（R37 教训） / set the truncation flag explicitly, lesson R37
    eErr   := 16#0001_0277; // 上溢码：超 255 已截断 / overflow code, truncated at the 255 cap
    bError     := TRUE; // 置错误标志 / raise error flag
    bValid     := FALSE; // 截断降级结果 / degraded truncated output
ELSE
    nUseB := nLenB; // 域内直通 / in-domain pass-through
END_IF

// 段 4｜复制 A 段：FOR 循环 + 255 越界 EXIT 守卫 / segment 4, copy the front part with the overrun guard
FOR nI := 1 TO nLenA DO
    IF nI > DL_CC_MAX THEN       (* 越界守卫（双重保险） EN: overrun guard *)
        EXIT;
    END_IF
    sResult[nI] := sA[nI]; // 逐字符复制 / char-by-char copy
END_FOR

// 段 5｜复制 B 段：目的位序 = A 段长加索引，超 255 即退出 / segment 5, copy the rear part, destination position = front length plus index
FOR nI := 1 TO nUseB DO
    IF (nLenA + nI) > DL_CC_MAX THEN   (* 越界守卫（双重保险） EN: overrun guard *)
        EXIT;
    END_IF
    sResult[nLenA + nI] := sB[nI]; // 逐字符复制 / char-by-char copy
END_FOR

// 段 6｜显式写终止符：总长未满 255 时在下一位置写空字符 / segment 6, write the terminator explicitly
IF nTotal < DL_CC_MAX THEN
    sResult[nTotal + 1] := '$00'; // 空字符终止符 / null terminator
END_IF
END_FUNCTION

(* ---- FC_DL_StringDeleteEx.st ---- *)
(*
    FC_DL_StringDeleteEx —— 删除指定区间防御包装（区间越界钳位，删除只缩不长）
    ------------------------------------------------------------------
    分类      : DL_MathData / String
    前缀      : FC_DL_
    版本      : 1.0.0
    溯源      : IEC 61131-3 标准语义的道莅防御性实现
                （内部委托平台内建函数，外围统一错误码/钳位/双语文档；
                  未复制任何闭源厂商源码，参考实现仅限 MIT/Apache 许可）
    平台      : 纯 IEC 61131-3，CODESYS / TwinCAT / InoProShop 通用
    作者      : 道莅代码库 · PLC编程专家（R15）
    ------------------------------------------------------------------
    功能说明  : 删除 sIn 自 nPos 位序（1 基）起的 nCount 个字符。删除只
                会缩短串长，结果恒不超 255，无截断标志需求。处理次序：
                ① 锁存源串长；② nCount <= 0 原样返回置 16#0001_01B5；③ nPos < 1
                钳 1 置 16#0001_01B3；④ nPos > len 原样返回置 16#0001_01B3；⑤ 区间尾
                nPos+nCount-1 > len 截到串尾置 16#0001_01B3（bValid=FALSE）；
                ⑥ 前段 + 后段逐字符复制（每轮 255 越界 EXIT 守卫），复制
                后显式写空字符终止符。返回值 TRUE 表示已执行完成。
    错误码    : 0000 正常 / 16#0001_01B3 入参越界（nPos 钳位/超长，区间尾截到串尾） / 16#0001_01B5 无效入参（nCount <= 0，原样返回）
    修订记录  : 2026-11-16 v1.0.0 首次入库（R15）
*)
FUNCTION FC_DL_StringDeleteEx : BOOL
VAR_INPUT
    sIn    : STRING(255); // 源串 [字符] / source string [chars]
    nPos   : INT; // 删除起始位序 [字符位序]，1 基 / delete start position [char position], 1-based
    nCount : INT; // 删除字符数 [字符]，<= 0 判无效 / char count to delete [chars], values at or below 0 invalid
END_VAR
VAR_OUTPUT
    sResult  : STRING(255); // 结果串 [字符] / result string [chars]
    eErr : UDINT; // 错误码，0=正常 / error id, 0=ok
    bError   : BOOL; // 是否出错，eErr 非 0 时为 TRUE / error flag, TRUE when eErr is nonzero
    bValid   : BOOL; // 输出是否有效可用 / output valid
END_VAR
VAR
    nI     : INT; // 循环索引 [字符位序]，1 基 / loop index [char position], 1-based
    nLen   : INT; // 锁存的源串有效长度 [字符] / latched effective source length [chars]
    nPosC  : INT; // 钳位后的删除起始位序 [字符位序] / clamped delete start position [char position]
    nEnd   : INT; // 删除区间尾位序 [字符位序]，已截到串尾 / delete end position, clipped to the string end [char position]
    nF     : INT; // 前段字符数 [字符] / front part char count [chars]
    nT     : INT; // 后段字符数 [字符] / rear part char count [chars]
END_VAR
VAR CONSTANT
    DL_DE_MAX : INT := 255; // 串型上限 [字符] / string type cap [chars]
END_VAR

// 段 1｜返回值与输出预置，任何早退路径不留脏码 / segment 1, preset return value and outputs
FC_DL_StringDeleteEx := TRUE; // 返回值预置 TRUE（已执行口径） / preset return to TRUE
sResult              := ''; // 结果串预置空串 / preset result to the empty string
eErr             := 16#0000_0000; // 错误码预置正常 / preset error id to ok
bError               := FALSE; // 错误标志预置无错 / preset error flag to FALSE
bValid               := TRUE; // 有效标志预置可用 / preset valid flag to TRUE

// 段 2｜源串有效长度一次锁存（空字符截止扫描 + 255 越界守卫） / segment 2, latch the effective source length once
nI   := 1; // 索引起始 [字符位序] / index start
nLen := 0; // 有效长度预置 [字符] / preset effective length
WHILE nI <= DL_DE_MAX DO
    IF nI > DL_DE_MAX THEN   (* 越界守卫（双重保险） EN: overrun guard *)
        EXIT;
    END_IF
    IF sIn[nI] = '$00' THEN  (* 首个空字符即串结束 EN: first null char ends the string *)
        EXIT;
    END_IF
    nLen := nI; // 记录最后非空位序 [字符] / record the last non-null position
    nI   := nI + 1; // 每轮自增 / per-iteration increment
END_WHILE

// 段 3｜无效入参闸：nCount <= 0 原样返回置 16#0001_01B5 / segment 3, invalid input gate, count at or below 0 returns the original with code 4
IF nCount <= 0 THEN
    FOR nI := 1 TO nLen DO
        IF nI > DL_DE_MAX THEN   (* 越界守卫（双重保险） EN: overrun guard *)
            EXIT;
        END_IF
        sResult[nI] := sIn[nI]; // 原样逐字符复制 / copy the original char by char
    END_FOR
    IF nLen < DL_DE_MAX THEN
        sResult[nLen + 1] := '$00'; // 空字符终止符 / null terminator
    END_IF
    eErr := 16#0001_01B5; // 无效入参码 / invalid input code
    bError   := TRUE; // 置错误标志 / raise error flag
    bValid   := FALSE; // 输出不可用 / output invalid
    RETURN;
END_IF

// 段 4｜位置钳位与越界组合闸：nPos < 1 钳 1；nPos > len 原样返回 / segment 4, position clamp and out-of-range combination gate
IF nPos < 1 THEN
    nPosC := 1; // 下越界钳 1 / clamped to 1
    eErr := 16#0001_01B3; // 入参越界码 / out-of-domain code
    bError := TRUE; // 置错误标志 / raise error flag
    bValid := FALSE; // 钳位降级 / degraded output
ELSE
    nPosC := nPos; // 域内直通 / in-domain pass-through
END_IF
IF nPosC > nLen THEN
    FOR nI := 1 TO nLen DO
        IF nI > DL_DE_MAX THEN   (* 越界守卫（双重保险） EN: overrun guard *)
            EXIT;
        END_IF
        sResult[nI] := sIn[nI]; // 起点超长原样返回 / start beyond length, original returned
    END_FOR
    IF nLen < DL_DE_MAX THEN
        sResult[nLen + 1] := '$00'; // 空字符终止符 / null terminator
    END_IF
    eErr := 16#0001_01B3; // 入参越界码（首事件优先不覆盖 16#0001_01B5） / out-of-domain code, first event kept
    bError   := TRUE; // 置错误标志 / raise error flag
    bValid   := FALSE; // 输出不可用 / output invalid
    RETURN;
END_IF

// 段 5｜区间尾截断闸：nPos+nCount-1 超 len 截到串尾置 16#0001_01B3 / segment 5, interval end clipping gate, end beyond the length clipped with code 1
nEnd := nPosC + nCount - 1; // 原始区间尾 [字符位序] / raw interval end
IF nEnd > nLen THEN
    nEnd := nLen; // 截到串尾 / clipped to the string end
    eErr := 16#0001_01B3; // 入参越界码 / out-of-domain code
    bError   := TRUE; // 置错误标志 / raise error flag
    bValid   := FALSE; // 区间被截短，输出降级 / interval clipped, degraded output
END_IF
nF := nPosC - 1; // 前段字符数 [字符] / front part char count
nT := nLen - nEnd; // 后段字符数 [字符] / rear part char count

// 段 6｜复制前段：FOR 循环 + 255 越界 EXIT 守卫 / segment 6, copy the front part with the overrun guard
FOR nI := 1 TO nF DO
    IF nI > DL_DE_MAX THEN       (* 越界守卫（双重保险） EN: overrun guard *)
        EXIT;
    END_IF
    sResult[nI] := sIn[nI]; // 逐字符复制 / char-by-char copy
END_FOR

// 段 7｜复制后段：源自 nEnd+1 起，目的位序顺延 / segment 7, copy the rear part
FOR nI := 1 TO nT DO
    IF (nF + nI) > DL_DE_MAX THEN    (* 目的侧越界守卫 EN: destination overrun guard *)
        EXIT;
    END_IF
    IF (nEnd + nI) > DL_DE_MAX THEN  (* 源侧越界守卫 EN: source overrun guard *)
        EXIT;
    END_IF
    sResult[nF + nI] := sIn[nEnd + nI]; // 逐字符复制 / char-by-char copy
END_FOR

// 段 8｜显式写终止符 / segment 8, write the terminator explicitly
IF (nF + nT) < DL_DE_MAX THEN
    sResult[nF + nT + 1] := '$00'; // 空字符终止符 / null terminator
END_IF
END_FUNCTION

(* ---- FC_DL_StringFindEx.st ---- *)
(*
    FC_DL_StringFindEx —— 子串查找防御包装（1 基返回位置，未找到不是错误）
    ------------------------------------------------------------------
    分类      : DL_MathData / String
    前缀      : FC_DL_
    版本      : 1.0.0
    溯源      : IEC 61131-3 标准语义的道莅防御性实现
                （内部委托平台内建函数，外围统一错误码/钳位/双语文档；
                  未复制任何闭源厂商源码，参考实现仅限 MIT/Apache 许可）
    平台      : 纯 IEC 61131-3，CODESYS / TwinCAT / InoProShop 通用
    作者      : 道莅代码库 · PLC编程专家（R15）
    ------------------------------------------------------------------
    功能说明  : 在 sHay 中自 nStart 位序（1 基）起查找 sNeedle 首次出现
                位置，返回 1 基位序；未找到返回 0 且 eErr=0000、
                bValid=TRUE（未找到不是错误）。sNeedle 为空串返回 0 置
                16#0001_01BA；nStart < 1 钳 1 置 16#0001_01B8；nStart > 主串长返回 0 置
                16#0001_01B8。双层循环：外层起点受 主串长-子串长+1 上限约束，
                内层匹配带 255 越界 EXIT 守卫，失配即断内层回退外层下一
                起点，无死循环风险。返回值即位置。
    错误码    : 0000 正常（含未找到返回 0） / 16#0001_01B8 入参越界（nStart 钳位或超主串长） / 16#0001_01BA 无效入参（sNeedle 为空串）
    修订记录  : 2026-11-16 v1.0.0 首次入库（R15）
*)
FUNCTION FC_DL_StringFindEx : INT
VAR_INPUT
    sHay    : STRING(255); // 主串 [字符] / haystack string [chars]
    sNeedle : STRING(255); // 子串 [字符] / needle string [chars]
    nStart  : INT; // 查找起始位序 [字符位序]，1 基 / search start position [char position], 1-based
END_VAR
VAR_OUTPUT
    eErr : UDINT; // 错误码，0=正常（含未找到） / error id, 0=ok including the not-found case
    bError   : BOOL; // 是否出错，eErr 非 0 时为 TRUE / error flag, TRUE when eErr is nonzero
    bValid   : BOOL; // 输出是否有效可用，未找到时保持 TRUE / output valid, stays TRUE for the not-found case
END_VAR
VAR
    nI       : INT; // 外层循环索引 [字符位序]，主串起点 / outer loop index [char position], haystack start
    nJ       : INT; // 内层循环索引 [字符位序]，子串偏移 / inner loop index [char position], needle offset
    nHayLen  : INT; // 锁存的主串有效长度 [字符] / latched effective haystack length [chars]
    nNeedLen : INT; // 锁存的子串有效长度 [字符] / latched effective needle length [chars]
    nStartC  : INT; // 钳位后的查找起点 [字符位序] / clamped search start [char position]
    nLimit   : INT; // 外层起点上限 [字符位序] / outer start upper bound [char position]
    bMatch   : BOOL; // 内层匹配成功标志 / inner-loop match success flag
END_VAR
VAR CONSTANT
    DL_FD_MAX : INT := 255; // 串型上限 [字符] / string type cap [chars]
END_VAR

// 段 1｜返回值与错误状态预置，任何早退路径不留脏码 / segment 1, preset return value and error states
FC_DL_StringFindEx := 0; // 返回值预置 0（未找到口径）[字符位序] / preset return to 0, not-found semantics
eErr           := 16#0000_0000; // 错误码预置正常 / preset error id to ok
bError             := FALSE; // 错误标志预置无错 / preset error flag to FALSE
bValid             := TRUE; // 有效标志预置可用（未找到也是有效结果） / preset valid to TRUE, not-found is a valid result

// 段 2｜两串有效长度各一次锁存（空字符截止扫描 + 255 越界守卫） / segment 2, latch both effective lengths once
nI       := 1; // 索引起始 [字符位序] / index start
nHayLen  := 0; // 主串长度预置 [字符] / preset haystack length
WHILE nI <= DL_FD_MAX DO
    IF nI > DL_FD_MAX THEN    (* 越界守卫（双重保险） EN: overrun guard *)
        EXIT;
    END_IF
    IF sHay[nI] = '$00' THEN  (* 首个空字符即串结束 EN: first null char ends the string *)
        EXIT;
    END_IF
    nHayLen := nI; // 记录主串最后非空位序 [字符] / record the last non-null position
    nI      := nI + 1; // 每轮自增 / per-iteration increment
END_WHILE
nI       := 1; // 索引复位 / reset index
nNeedLen := 0; // 子串长度预置 [字符] / preset needle length
WHILE nI <= DL_FD_MAX DO
    IF nI > DL_FD_MAX THEN    (* 越界守卫（双重保险） EN: overrun guard *)
        EXIT;
    END_IF
    IF sNeedle[nI] = '$00' THEN (* 首个空字符即串结束 EN: first null char ends the string *)
        EXIT;
    END_IF
    nNeedLen := nI; // 记录子串最后非空位序 [字符] / record the last non-null position
    nI       := nI + 1; // 每轮自增 / per-iteration increment
END_WHILE

// 段 3｜无效入参闸：子串空串返回 0 置 16#0001_01BA / segment 3, invalid input gate, empty needle returns 0 with code 4
IF nNeedLen <= 0 THEN
    eErr := 16#0001_01BA; // 无效入参码 / invalid input code
    bError   := TRUE; // 置错误标志 / raise error flag
    bValid   := FALSE; // 输出不可用 / output invalid
    RETURN;
END_IF

// 段 4｜起点钳位闸：nStart < 1 钳 1 置 16#0001_01B8；nStart > 主串长返回 0 置 16#0001_01B8 / segment 4, start clamp gate
IF nStart < 1 THEN
    nStartC := 1; // 下越界钳 1 / clamped to 1
    eErr := 16#0001_01B8; // 入参越界码 / out-of-domain code
    bError   := TRUE; // 置错误标志 / raise error flag
    bValid   := FALSE; // 钳位降级 / degraded output
ELSE
    nStartC := nStart; // 域内直通 / in-domain pass-through
END_IF
IF nStartC > nHayLen THEN
    FC_DL_StringFindEx := 0; // 起点超主串长返回 0 / start beyond haystack length returns 0
    eErr := 16#0001_01B8; // 入参越界码 / out-of-domain code
    bError   := TRUE; // 置错误标志 / raise error flag
    bValid   := FALSE; // 输出不可用 / output invalid
    RETURN;
END_IF

// 段 5｜双层查找：外层起点上限 = 主串长减子串长加一，内层失配即断回退外层 / segment 5, two-layer search, outer bounded by haystack minus needle plus one, inner breaks on mismatch
nLimit := nHayLen - nNeedLen + 1; // 外层起点上限 [字符位序] / outer start upper bound
FOR nI := nStartC TO nLimit DO
    bMatch := TRUE; // 匹配标志预置成功 / preset the match flag to success
    nJ := 1; // 内层索引起始 [字符位序] / inner index start
    WHILE nJ <= nNeedLen DO
        IF (nI + nJ - 1) > DL_FD_MAX THEN    (* 主串侧越界守卫（双重保险） EN: haystack overrun guard *)
            bMatch := FALSE; // 越界即失配 / overrun means mismatch
            EXIT; // 断内层回退外层 / break the inner loop
        END_IF
        IF sHay[nI + nJ - 1] <> sNeedle[nJ] THEN   (* 逐字符比对 EN: char-by-char compare *)
            bMatch := FALSE; // 失配 / mismatch
            EXIT; // 断内层回退外层下一起点，无死循环 / break the inner loop, outer advances, no hang
        END_IF
        nJ := nJ + 1; // 内层自增 / inner increment
    END_WHILE
    IF bMatch THEN
        FC_DL_StringFindEx := nI; // 命中返回 1 基位置 / hit, return the 1-based position
        RETURN;
    END_IF
END_FOR

// 段 6｜未找到收口：返回预置 0，错误码保持 0000，bValid 保持 TRUE / segment 6, not-found closure, return the preset 0 with no error
END_FUNCTION

(* ---- FC_DL_StringInsertEx.st ---- *)
(*
    FC_DL_StringInsertEx —— 指定位置插入防御包装（位置钳位 + 255 截断显式置标志）
    ------------------------------------------------------------------
    分类      : DL_MathData / String
    前缀      : FC_DL_
    版本      : 1.0.0
    溯源      : IEC 61131-3 标准语义的道莅防御性实现
                （内部委托平台内建函数，外围统一错误码/钳位/双语文档；
                  未复制任何闭源厂商源码，参考实现仅限 MIT/Apache 许可）
    平台      : 纯 IEC 61131-3，CODESYS / TwinCAT / InoProShop 通用
    作者      : 道莅代码库 · PLC编程专家（R15）
    ------------------------------------------------------------------
    功能说明  : 在 sIn 的 nPos 位序（1 基）前插入 sIns，插入后 sIns 首字
                符位于 nPos 处。处理次序写死：① 锁存源串/插入串长度；
                ② 位置钳位：nPos < 1 钳 1、nPos > len+1 钳 len+1，置 16#0001_01AE；
                ③ 前段/插入段/后段三段配额预分配，插入段配额 = 255 - 前
                段长 - 后段长，超配额时按 R37 范式先置 bTruncated=TRUE 与
                16#0001_027C 再截断；④ 逐字符三段复制，每轮带 255 越界 EXIT 守卫，
                复制后显式写空字符终止符。返回值 TRUE 表示已执行完成。
    错误码    : 0000 正常 / 16#0001_01AE 入参越界（nPos 已钳位） / 16#0001_027C 上溢下溢（结果超 255，已显式截断，bTruncated=TRUE）
    修订记录  : 2026-11-16 v1.0.0 首次入库（R15）
*)
FUNCTION FC_DL_StringInsertEx : BOOL
VAR_INPUT
    sIn  : STRING(255); // 源串 [字符] / source string [chars]
    sIns : STRING(255); // 插入串 [字符] / string to insert [chars]
    nPos : INT; // 插入位序 [字符位序]，1 基，插入后 sIns 首字符居此 / insert position [char position], 1-based, first inserted char lands here
END_VAR
VAR_OUTPUT
    sResult    : STRING(255); // 结果串 [字符] / result string [chars]
    eErr : UDINT; // 错误码，0=正常，1=位置钳位，2=超 255 截断 / error id, 0=ok, 1=position clamped, 2=explicit truncation at the 255 cap
    bError     : BOOL; // 是否出错，eErr 非 0 时为 TRUE / error flag, TRUE when eErr is nonzero
    bValid     : BOOL; // 输出是否有效可用 / output valid
    bTruncated : BOOL; // 截断标志，发生 255 截断时 TRUE（R37 范式） / truncation flag, TRUE when the 255 cap truncated content
END_VAR
VAR
    nI       : INT; // 循环索引 [字符位序]，1 基 / loop index [char position], 1-based
    nLen     : INT; // 锁存的源串有效长度 [字符] / latched effective source length [chars]
    nInsLen  : INT; // 锁存的插入串有效长度 [字符] / latched effective insert length [chars]
    nPosC    : INT; // 钳位后的插入位序 [字符位序] / clamped insert position [char position]
    nF       : INT; // 前段字符数 [字符]，nPos 减一 / front part char count [chars]
    nT       : INT; // 后段字符数 [字符] / rear part char count [chars]
    nInsUse  : INT; // 插入段实际复制数 [字符]，受 255 配额钳制 / chars actually copied from the insert [chars]
    nTot     : INT; // 结果总长 [字符] / total result length [chars]
END_VAR
VAR CONSTANT
    DL_IN_MAX : INT := 255; // 串型上限 [字符] / string type cap [chars]
END_VAR

// 段 1｜返回值与输出预置，任何早退路径不留脏码 / segment 1, preset return value and outputs
FC_DL_StringInsertEx := TRUE; // 返回值预置 TRUE（已执行口径） / preset return to TRUE
sResult              := ''; // 结果串预置空串 / preset result to the empty string
eErr             := 16#0000_0000; // 错误码预置正常 / preset error id to ok
bError               := FALSE; // 错误标志预置无错 / preset error flag to FALSE
bValid               := TRUE; // 有效标志预置可用 / preset valid flag to TRUE
bTruncated           := FALSE; // 截断标志预置无截断 / preset truncation flag to FALSE

// 段 2｜两串有效长度各一次锁存（空字符截止扫描 + 255 越界守卫） / segment 2, latch both effective lengths once
nI      := 1; // 索引起始 [字符位序] / index start
nLen    := 0; // 源串长度预置 [字符] / preset source length
WHILE nI <= DL_IN_MAX DO
    IF nI > DL_IN_MAX THEN    (* 越界守卫（双重保险） EN: overrun guard *)
        EXIT;
    END_IF
    IF sIn[nI] = '$00' THEN   (* 首个空字符即串结束 EN: first null char ends the string *)
        EXIT;
    END_IF
    nLen := nI; // 记录源串最后非空位序 [字符] / record the last non-null position
    nI   := nI + 1; // 每轮自增 / per-iteration increment
END_WHILE
nI      := 1; // 索引复位 / reset index
nInsLen := 0; // 插入串长度预置 [字符] / preset insert length
WHILE nI <= DL_IN_MAX DO
    IF nI > DL_IN_MAX THEN    (* 越界守卫（双重保险） EN: overrun guard *)
        EXIT;
    END_IF
    IF sIns[nI] = '$00' THEN  (* 首个空字符即串结束 EN: first null char ends the string *)
        EXIT;
    END_IF
    nInsLen := nI; // 记录插入串最后非空位序 [字符] / record the last non-null position
    nI      := nI + 1; // 每轮自增 / per-iteration increment
END_WHILE

// 段 3｜位置钳位闸：nPos < 1 钳 1，nPos > len+1 钳 len+1，置 16#0001_01AE / segment 3, position clamp gate, below 1 clamped to 1, beyond len plus 1 clamped to len plus 1, code 1
IF nPos < 1 THEN
    nPosC    := 1; // 下越界钳 1 / clamped to 1
    eErr := 16#0001_01AE; // 入参越界码 / out-of-domain code
    bError   := TRUE; // 置错误标志 / raise error flag
    bValid   := FALSE; // 钳位降级 / degraded output
ELSIF nPos > (nLen + 1) THEN
    nPosC    := nLen + 1; // 上越界钳到串尾后一位 / clamped to one past the end
    eErr := 16#0001_01AE; // 入参越界码 / out-of-domain code
    bError   := TRUE; // 置错误标志 / raise error flag
    bValid   := FALSE; // 钳位降级 / degraded output
ELSE
    nPosC := nPos; // 域内直通 / in-domain pass-through
END_IF
nF := nPosC - 1; // 前段字符数 [字符] / front part char count
nT := nLen - nF; // 后段字符数 [字符] / rear part char count

// 段 4｜插入段配额闸（R37 范式：先判定后写入，严禁静默回夹） / segment 4, insert quota gate, R37 paradigm, decide before writing
IF nInsLen > (DL_IN_MAX - nF - nT) THEN
    nInsUse := DL_IN_MAX - nF - nT; // 插入段配额，可为 0 / insert quota, may be zero
    bTruncated := TRUE; // 显式置截断标志（R37 教训） / set the truncation flag explicitly
    eErr   := 16#0001_027C; // 上溢码：超 255 已截断 / overflow code, truncated
    bError     := TRUE; // 置错误标志 / raise error flag
    bValid     := FALSE; // 截断降级结果 / degraded truncated output
ELSE
    nInsUse := nInsLen; // 域内直通 / in-domain pass-through
END_IF

// 段 5｜复制前段：FOR 循环 + 255 越界 EXIT 守卫 / segment 5, copy the front part with the overrun guard
FOR nI := 1 TO nF DO
    IF nI > DL_IN_MAX THEN        (* 越界守卫（双重保险） EN: overrun guard *)
        EXIT;
    END_IF
    sResult[nI] := sIn[nI]; // 逐字符复制 / char-by-char copy
END_FOR

// 段 6｜复制插入段：目的位序 = 前段长加索引，超 255 即退出 / segment 6, copy the insert part
FOR nI := 1 TO nInsUse DO
    IF (nF + nI) > DL_IN_MAX THEN     (* 越界守卫（双重保险） EN: overrun guard *)
        EXIT;
    END_IF
    sResult[nF + nI] := sIns[nI]; // 逐字符复制 / char-by-char copy
END_FOR

// 段 7｜复制后段：源 sIn 自 nF+1 起，目的位序顺延 / segment 7, copy the rear part from the source
FOR nI := 1 TO nT DO
    IF (nF + nInsUse + nI) > DL_IN_MAX THEN   (* 越界守卫（双重保险） EN: overrun guard *)
        EXIT;
    END_IF
    IF (nF + nI) > DL_IN_MAX THEN             (* 源侧越界守卫 EN: source overrun guard *)
        EXIT;
    END_IF
    sResult[nF + nInsUse + nI] := sIn[nF + nI]; // 逐字符复制 / char-by-char copy
END_FOR

// 段 8｜显式写终止符 / segment 8, write the terminator explicitly
nTot := nF + nInsUse + nT; // 结果总长 [字符] / total result length
IF nTot < DL_IN_MAX THEN
    sResult[nTot + 1] := '$00'; // 空字符终止符 / null terminator
END_IF
END_FUNCTION

(* ---- FC_DL_StringLeftEx.st ---- *)
(*
    FC_DL_StringLeftEx —— 取左 n 字符防御包装（n 越界钳位 + 255 守卫逐字符复制）
    ------------------------------------------------------------------
    分类      : DL_MathData / String
    前缀      : FC_DL_
    版本      : 1.0.0
    溯源      : IEC 61131-3 标准语义的道莅防御性实现
                （内部委托平台内建函数，外围统一错误码/钳位/双语文档；
                  未复制任何闭源厂商源码，参考实现仅限 MIT/Apache 许可）
    平台      : 纯 IEC 61131-3，CODESYS / TwinCAT / InoProShop 通用
    作者      : 道莅代码库 · PLC编程专家（R15）
    ------------------------------------------------------------------
    功能说明  : 取源串左侧 nCount 个字符到 sResult。采用逐字符 FOR 复制
                （跨平台口径，不依赖平台 LEFT 行为差异），每轮带 255 越
                界 EXIT 守卫，复制后显式写空字符终止符。nCount <= 0 返回
                空串置 16#0001_01A1；nCount > 实际长度返回全串并置 16#0001_019F（bValid=
                FALSE，截断诉求由错误码显式体现）。返回值 TRUE 表示函数
                已执行完成，结果总在 sResult 中，错误详情经 eErr 传递。
    错误码    : 0000 正常 / 16#0001_019F 入参越界（nCount 超实际长度，已返回全串） / 16#0001_01A1 无效入参（nCount <= 0）
    修订记录  : 2026-11-16 v1.0.0 首次入库（R15）
*)
FUNCTION FC_DL_StringLeftEx : BOOL
VAR_INPUT
    sIn    : STRING(255); // 源串 [字符] / source string [chars]
    nCount : INT; // 请求取左字符数 [字符]，<= 0 判无效 / requested left char count [chars], values at or below 0 invalid
END_VAR
VAR_OUTPUT
    sResult  : STRING(255); // 结果串 [字符]，左 nCount 字符 / result string [chars], left nCount chars
    eErr : UDINT; // 错误码，0=正常 / error id, 0=ok
    bError   : BOOL; // 是否出错，eErr 非 0 时为 TRUE / error flag, TRUE when eErr is nonzero
    bValid   : BOOL; // 输出是否有效可用 / output valid
END_VAR
VAR
    nI   : INT; // 循环索引 [字符位序]，1 基 / loop index [char position], 1-based
    nLen : INT; // 锁存的源串有效长度 [字符] / latched effective source length [chars]
    nUse : INT; // 实际复制字符数 [字符] / chars actually copied [chars]
END_VAR
VAR CONSTANT
    DL_LF_MAX : INT := 255; // 串型上限 [字符] / string type cap [chars]
END_VAR

// 段 1｜返回值与输出预置，任何早退路径不留脏码 / segment 1, preset return value and outputs so no early exit leaves stale states
FC_DL_StringLeftEx := TRUE; // 返回值预置 TRUE（已执行口径） / preset return to TRUE, executed semantics
sResult            := ''; // 结果串预置空串 / preset result to the empty string
eErr           := 16#0000_0000; // 错误码预置正常 / preset error id to ok
bError             := FALSE; // 错误标志预置无错 / preset error flag to FALSE
bValid             := TRUE; // 有效标志预置可用 / preset valid flag to TRUE

// 段 2｜源串有效长度一次锁存（空字符截止扫描 + 255 越界守卫） / segment 2, latch the effective source length once with the null-terminated scan and overrun guard
nI   := 1; // 索引起始 [字符位序] / index start
nLen := 0; // 有效长度预置 [字符] / preset effective length
WHILE nI <= DL_LF_MAX DO
    IF nI > DL_LF_MAX THEN   (* 越界守卫（双重保险） EN: overrun guard, defense in depth *)
        EXIT;
    END_IF
    IF sIn[nI] = '$00' THEN  (* 首个空字符即串结束 EN: first null character marks the string end *)
        EXIT;
    END_IF
    nLen := nI; // 记录最后非空字符位序 [字符] / record the last non-null char position
    nI   := nI + 1; // 每轮自增 / per-iteration increment
END_WHILE

// 段 3｜入参域闸门：nCount <= 0 无效置 16#0001_01A1；nCount 超长度钳到全长置 16#0001_019F / segment 3, input domain gate, count at or below 0 invalid with code 4, count beyond length clamped to full length with code 1
IF nCount <= 0 THEN
    sResult  := ''; // 无效入参返回空串 / invalid input returns the empty string
    eErr := 16#0001_01A1; // 无效入参码 / invalid input code
    bError   := TRUE; // 置错误标志 / raise error flag
    bValid   := FALSE; // 输出不可用 / output invalid
    RETURN;
ELSIF nCount > nLen THEN
    nUse    := nLen; // 请求超长，钳到全串长 / request beyond length, clamped to full length
    eErr := 16#0001_019F; // 入参越界码：截断诉求显式置码 / out-of-domain code, truncation intent made explicit
    bError   := TRUE; // 置错误标志 / raise error flag
    bValid   := FALSE; // 输出为截断降级结果 / output is a degraded truncated result
ELSE
    nUse := nCount; // 域内直通 / in-domain pass-through
END_IF

// 段 4｜逐字符复制（跨平台口径）：FOR 循环 + 255 越界 EXIT 守卫 / segment 4, char-by-char copy for cross-platform portability, for loop with the 255 overrun EXIT guard
FOR nI := 1 TO nUse DO
    IF nI > DL_LF_MAX THEN       (* 越界守卫（双重保险） EN: overrun guard, defense in depth *)
        EXIT;
    END_IF
    sResult[nI] := sIn[nI]; // 逐字符复制 / char-by-char copy
END_FOR

// 段 5｜显式写终止符：nUse 未满 255 时在下一位置写空字符 / segment 5, write the terminator explicitly, at the next position when nUse is below the cap
IF nUse < DL_LF_MAX THEN
    sResult[nUse + 1] := '$00'; // 空字符终止符 / null terminator
END_IF
END_FUNCTION

(* ---- FC_DL_StringLenEx.st ---- *)
(*
    FC_DL_StringLenEx —— 字符串有效长度防御包装（空字符截止 + 尾空格可选回退）
    ------------------------------------------------------------------
    分类      : DL_MathData / String
    前缀      : FC_DL_
    版本      : 1.0.0
    溯源      : IEC 61131-3 标准语义的道莅防御性实现
                （内部委托平台内建函数，外围统一错误码/钳位/双语文档；
                  未复制任何闭源厂商源码，参考实现仅限 MIT/Apache 许可）
    平台      : 纯 IEC 61131-3，CODESYS / TwinCAT / InoProShop 通用
    作者      : 道莅代码库 · PLC编程专家（R15）
    ------------------------------------------------------------------
    功能说明  : 返回输入字符串的有效长度。自位序 1 扫描至 255，遇第一个
                空字符即截止（长度取最后非空字符位序）；随后按入参
                bTrimTrailingSpace 决定是否回退尾部空格（TRUE 回退、FALSE
                计入）。WHILE 循环每轮带 255 越界 EXIT 守卫，空格回退循环
                用嵌套 IF 结构避免对短路求值的依赖。长度 0 为正常结果
                （eErr=0000、bValid=TRUE），不置任何错误码。
    错误码    : 0000 正常（含空串长度 0 的正常输出）
    修订记录  : 2026-11-16 v1.0.0 首次入库（R15）
*)
FUNCTION FC_DL_StringLenEx : INT
VAR_INPUT
    sIn                : STRING(255); // 输入字符串 [字符] / input string [chars]
    bTrimTrailingSpace : BOOL; // TRUE=尾部空格不计入长度，FALSE=尾部空格计入 / TRUE=trailing spaces not counted, FALSE=trailing spaces counted
END_VAR
VAR_OUTPUT
    eErr : UDINT; // 错误码，本件仅 0=正常 / error id, this unit only 0=ok
    bError   : BOOL; // 是否出错，eErr 非 0 时为 TRUE / error flag, TRUE when eErr is nonzero
    bValid   : BOOL; // 输出是否有效可用 / output valid
END_VAR
VAR
    nI   : INT; // 循环索引 [字符位序]，1 基 / loop index [char position], 1-based
    nLen : INT; // 有效长度 [字符]，最后非空字符位序 / effective length [chars], position of the last non-null char
END_VAR
VAR CONSTANT
    DL_SL_MAX : INT := 255; // 串型上限 [字符]，定长 STRING 的隐式容量 / string type cap [chars], implicit capacity of a fixed-length STRING
END_VAR

// 段 1｜返回值与错误状态预置，任何早退路径不留脏码 / segment 1, preset return value and error states
FC_DL_StringLenEx := 0; // 返回值预置 0 [字符] / preset return to 0
eErr          := 16#0000_0000; // 错误码预置正常 / preset error id to ok
bError            := FALSE; // 错误标志预置无错 / preset error flag to FALSE
bValid            := TRUE; // 有效标志预置可用 / preset valid flag to TRUE

// 段 2｜空字符截止扫描：WHILE 循环 + 每轮自增 + 255 越界 EXIT 守卫 / segment 2, null-terminated scan, while loop with per-iteration increment and the 255 overrun EXIT guard
nI   := 1; // 索引自位序 1 起始 [字符位序] / index starts at position 1
nLen := 0; // 有效长度预置 0（空串口径）[字符] / preset effective length to 0 for the empty-string case
WHILE nI <= DL_SL_MAX DO
    IF nI > DL_SL_MAX THEN   (* 越界守卫（双重保险，严禁越界索引） EN: overrun guard, defense in depth, no out-of-bound indexing *)
        EXIT;
    END_IF
    IF sIn[nI] = '$00' THEN  (* 首个空字符即串结束 EN: first null character marks the string end *)
        EXIT;
    END_IF
    nLen := nI; // 记录最后非空字符位序 [字符] / record the last non-null char position
    nI   := nI + 1; // 每轮自增 [字符位序] / per-iteration increment
END_WHILE

// 段 3｜尾部空格回退（可选）：嵌套 IF 结构，不依赖短路求值，nLen=0 时安全终止 / segment 3, optional trailing space trim, nested-if structure without short-circuit reliance, safe at zero length
IF bTrimTrailingSpace THEN
    WHILE nLen > 0 DO
        IF sIn[nLen] = ' ' THEN
            nLen := nLen - 1; // 尾部空格回退一格 [字符] / trim one trailing space
        ELSE
            EXIT; // 非空格字符，回退结束 / non-space char reached, trimming done
        END_IF
    END_WHILE
END_IF

// 段 4｜输出有效长度 / segment 4, output the effective length
FC_DL_StringLenEx := nLen; // 输出有效长度 [字符] / output the effective length
END_FUNCTION

(* ---- FC_DL_StringMidEx.st ---- *)
(*==============================================================================
 * 组件名称 (Component)  : FC_DL_StringMidEx
 * 所属子库 (Sublibrary) : DL_MathData
 * 当前版本 (Version)    : 1.0.0
 * 兼容性   (Platform)   : CODESYS 3.5 / TwinCAT 3 / 汇川 InoProShop / Machine Expert
 *                         仅依赖 Standard.library 的 MID / LEN / MIN 内建函数，
 *                         不重实现取子串内核，无厂商字符串方言依赖
 * 功能一句话 (Summary)  : MID 取子串防御包装：起点/长度域闸门钳位 +
 *                         255 上限截断显式置标志（R37 教训：严禁静默回夹）。
 * 功能描述 (Function)   : 从源串 sIn 的 iStart 位序（1 基）起取 iLen 个字符。
 *                         处理次序写死（R37 范式「先判定后写入」）：
 *                         ① LEN 一次锁存源串长（防调用中串被改写的时序歧义）；
 *                         ② 参数域闸门——iStart < 1 钳 1、iLen < 0 钳 0，
 *                         置信息码；③ 越界组合闸——起点超串长返回空串置码；
 *                         ④ 255 上限截断闸——请求长度超串型上限先置截断
 *                         标志再钳长，最后才委托内建 MID，杜绝静默回夹。
 * 溯源     (Origin)     : IEC 61131-3 标准语义的道莅防御性实现
 *                         （接口语义由 IEC 61131-3 定义，clean-room 重写，
 *                         参考公开标准条款）
 * 码位     (Diag Codes) : 信息级 16#0001_015C（本件独占）：
 *                           参数钳位（iStart<1 钳 1 / iLen<0 钳 0）或起点
 *                           超出串长（含空串输入，返回空串）；
 *                         信息级 16#0001_015D（本件独占）：
 *                           请求子串超串型上限 255，已显式截断（R37 教训：
 *                           定长串截断必须显式置位，严禁静默回夹）。
 * 类型裁定 (Type Note)  : 码位段 16#0001_xxxx 为全库共享 32 位段，WORD 容量不足，
 *                         故 eErr 采用 UDINT 承载（与库内 uErrorId : UDINT 惯例
 *                         一致，沿 R14 批 3 同一裁定）。
 * 依赖     (Depends)    : 无 DL_ 内部依赖；Standard.library: MID / LEN / MIN
 * 红线自检 (Redline)    : R1 ✓ 零全局变量与外部变量引用 ｜ R2 ✓ 零物理 IO 地址直写
 *                         R3 ✓ 纯 IEC 61131-3 ｜ R4 ✓ 域闸门先行 + 截断先置标志后钳长
 *                         R5 ✓ 全变量中英双语同行注释
 *                         R6 N/A（纯函数，无 CASE/ENUM 状态机，按批 4 口径标 N/A）
 *                         R7 N/A（FC 为纯函数，无实例调用，头注释显式说明）
 * 防御行为声明 (Defense): ① 处理次序写死「锁存 → 钳位 → 越界闸 → 截断闸 →
 *                           委托内建」，截断判定先于任何写入（R37 范式，
 *                           与库内样板件 FC_DL_StringFixedField 同源）；
 *                         ② LEN 只调用一次锁存到局部变量，后续边界全部用
 *                           锁存值判定——调用拍内源串再被改写也不产生
 *                           「边界用旧长、切片用新长」的时序歧义；
 *                         ③ iStart < 1 钳 1、iLen < 0 钳 0：钳位是正常防御
 *                           行为，置信息码不置故障码；
 *                         ④ 起点超串长（含空串）返回空串并置信息码，
 *                           不调用内建 MID（部分平台对越界起点行为不一）；
 *                         ⑤ 请求长度先按可用串长取 MIN，再对串型上限 255
 *                           截断：超限先置截断标志 16#0001_015D，再钳到 255
 *                           委托内建——MID 的静默回夹绝不作为唯一防线；
 *                         ⑥ 首事件优先：多条件同拍命中时保留先置的码，
 *                           后续码不覆盖，便于现场定位第一诱因；
 *                         ⑦ 串型上限 255 提为只读常量，禁魔法数。
 * 修订历史 (Revision)   :
 *   2026-11-16  v1.0.0  首版入库（R14 批 4 · T0 快车道）
 *============================================================================*)
FUNCTION FC_DL_StringMidEx : STRING
VAR_INPUT
    sIn    : STRING; // 源串 [字符]，定长串型，上限 255 / Source string [chars], fixed-length type, cap 255
    iStart : INT;    // 起始位序 [字符]，1 基，< 1 钳 1 / Start position [chars], 1-based, values below 1 clamped to 1
    iLen   : INT;    // 取长 [字符]，< 0 钳 0 / Length to extract [chars], values below 0 clamped to 0
END_VAR
VAR_OUTPUT
    eErr : UDINT; // 错误码，16#0001_015C=参数钳位或起点越界，16#0001_015D=超 255 显式截断，0=无事件 / Error code, 16#0001_015C=parameter clamped or start beyond length, 16#0001_015D=explicit truncation at the 255 cap, 0=no event
END_VAR
VAR
    nSrcLen : INT; // 锁存的源串长 [字符]，LEN 只调用一次 / Latched source length [chars], LEN called exactly once
    nPos    : INT; // 钳位后起始位序 [字符]，域 >= 1 / Clamped start position [chars], domain >= 1
    nLenC   : INT; // 钳位后取长 [字符]，域 >= 0 / Clamped extraction length [chars], domain >= 0
    nAvail  : INT; // 自起点起可用字符数 [字符] / Characters available from the start position [chars]
    nReq    : INT; // 请求取长 [字符]，取长与可用长取小 / Requested length [chars], min of clamped length and available length
    nUse    : INT; // 实际委托取长 [字符]，域 0 到 255 / Length actually delegated [chars], range 0 to 255
END_VAR
VAR CONSTANT
    DL_SM_MAX : INT := 255; // 串型上限 [字符]，定长 STRING 的隐式容量 / String type cap [chars], implicit capacity of a fixed-length STRING
END_VAR

(*------------------------------------------------------------------------------
 * 段 1｜返回值与错误码预置：先归零，任何早退路径都不会留下脏码
 *      Preset return value and error code so no early-exit path leaves a stale code
 *-----------------------------------------------------------------------------*)
FC_DL_StringMidEx := '';          // 返回值预置空串 [字符] / Preset return value to the empty string
eErr              := 16#0000_0000;   // 错误码预置无事件 / Preset error code to no event

(*------------------------------------------------------------------------------
 * 段 2｜源串长一次锁存（防御声明②）：后续边界全部用锁存值，
 *      消灭「边界用旧长、切片用新长」的时序歧义
 *      Latch the source length once (defense note 2): all bounds use the
 *      latched value, eliminating stale-length versus fresh-slice races
 *-----------------------------------------------------------------------------*)
nSrcLen := LEN(sIn);   // LEN 一次锁存 [字符] / Latch LEN exactly once [chars]

(*------------------------------------------------------------------------------
 * 段 3｜参数域闸门（防御声明③）：iStart < 1 钳 1、iLen < 0 钳 0，
 *      置信息码（首事件优先，防御声明⑥）
 *      Parameter domain gate (defense note 3): iStart below 1 clamped to 1,
 *      iLen below 0 clamped to 0, informational code raised (first-event
 *      priority per defense note 6)
 *-----------------------------------------------------------------------------*)
IF iStart < 1 THEN
    nPos := 1;              // 起始位序钳 1 [字符] / Start position clamped to 1 [chars]
    eErr := 16#0001_015C;   // 信息码：起始位序越下界已钳位 / Informational: start position below the lower bound, clamped
ELSE
    nPos := iStart;         // 域内直通 [字符] / In-domain pass-through [chars]
END_IF

IF iLen < 0 THEN
    nLenC := 0;             // 取长钳 0（空串结果）[字符] / Length clamped to 0 (empty result) [chars]
    IF eErr = 16#0000_0000 THEN
        eErr := 16#0001_015C;   // 信息码：取长越下界已钳位（首事件优先不覆盖）/ Informational: length below the lower bound, clamped (first event kept)
    END_IF
ELSE
    nLenC := iLen;          // 域内直通 [字符] / In-domain pass-through [chars]
END_IF

(*------------------------------------------------------------------------------
 * 段 4｜越界组合闸（防御声明④）：起点超锁存串长（含空串输入）返回空串，
 *      不调用内建 MID（平台对越界起点行为不一）
 *      Out-of-range combination gate (defense note 4): start beyond the latched
 *      length (including an empty input) returns the empty string without
 *      calling the built-in MID (platform behavior differs on bad starts)
 *-----------------------------------------------------------------------------*)
IF nPos > nSrcLen THEN
    FC_DL_StringMidEx := '';   // 起点越界返回空串 [字符] / Start beyond length, empty string returned
    IF eErr = 16#0000_0000 THEN
        eErr := 16#0001_015C;   // 信息码：起点超出串长（空串输入同此码）/ Informational: start beyond the string length (empty input shares this code)
    END_IF
    RETURN;                    // 早退，不进内建 / Early exit, built-in not called
END_IF

(*------------------------------------------------------------------------------
 * 段 5｜截断闸（防御声明①⑤⑦）：先按可用长取 MIN，再对 255 上限判定——
 *      超限先置截断标志，后钳长，最后才写结果（R37 范式：先判定后写入）
 *      Truncation gate (defense notes 1, 5 and 7): MIN against the available
 *      length first, then judge the 255 cap — set the truncation flag before
 *      clamping, write the result last (R37 paradigm: decide before writing)
 *-----------------------------------------------------------------------------*)
nAvail := nSrcLen - nPos + 1;   // 自起点起可用字符数 [字符] / Characters available from the start [chars]
nReq   := MIN(nLenC, nAvail);   // 请求取长 = 钳位取长与可用长取小 [字符] / Requested length, min of clamped and available [chars]

IF nReq > DL_SM_MAX THEN
    nUse := DL_SM_MAX;          // 请求超 255，钳到串型上限 [字符] / Request beyond 255, clamped to the string cap [chars]
    IF eErr = 16#0000_0000 THEN
        eErr := 16#0001_015D;   // 信息码：超 255 显式截断（严禁静默回夹，R37 教训）/ Informational: explicit truncation at the 255 cap (silent clipping forbidden, lesson R37)
    END_IF
ELSIF nReq <= 0 THEN
    nUse := 0;                  // 取长为 0，空串结果 [字符] / Zero length, empty result [chars]
ELSE
    nUse := nReq;               // 域内直通 [字符] / In-domain pass-through [chars]
END_IF

(*------------------------------------------------------------------------------
 * 段 6｜委托内建内核（防御声明⑤）：nUse 已锁死在 0 到 255 安全域，
 *      nPos 已锁死在 1 到锁存串长域，MID 无越界可能
 *      Delegation to the built-in kernel (defense note 5): nUse locked in
 *      0 to 255, nPos locked in 1 to the latched length, MID cannot overrun
 *-----------------------------------------------------------------------------*)
IF nUse = 0 THEN
    FC_DL_StringMidEx := '';   // 零长请求直接空串返回 [字符] / Zero-length request returns the empty string
ELSE
    FC_DL_StringMidEx := MID(sIn, nUse, nPos);   // 委托内建 MID 内核，不自实现切片 / Delegate to the built-in MID kernel, no re-implementation
END_IF
END_FUNCTION

(* ---- FC_DL_StringPad.st ---- *)
(*==============================================================================
 * 组件名称 (Component)  : FC_DL_StringPad
 * 溯源说明 (Provenance) : IEC 61131-3 标准语义的道莅防御性实现（零检索变体线）
 * 所属子库 (Sublibrary) : DL_MathData / StringOps
 * 当前版本 (Version)    : 1.0.0
 * 兼容性   (Platform)   : CODESYS 3.5 / TwinCAT 3 / 汇川 InoProShop；
 *                         纯 IEC 61131-3（第 3 版），仅用标准字符串函数 LEN/CONCAT
 * 组件分类 (Category)   : 函数（TYPE E_DL_PadSide :
(
    eLeft   := 0, // 左填充 / Left padding
    eRight  := 1, // 右填充 / Right padding
    eCenter := 2  // 居中填充 / Center padding
);
END_TYPE

FUNCTION）· 字符串定长填充（无状态纯函数）
 * 功能一句话 (Summary)  : 左/右/居中填充至目标长度；越界显式截断并置标志。
 * 边界与安全 (Boundary) : ①目标长度大于 255 → 钳 255 并置 bTruncated；
 *                         ②源串超长按目标长度截断并置 bTruncated（禁静默回夹）；
 *                         ③填充字符取首字符，空串降级为空格并置信息码；
 *                         ④居中奇偶差一优先填左侧（规格验收向量 ③）；
 *                         ⑤非法枚举侧别按右填充防御降级（03C2 保留不赋值）；
 *                         ⑥纯函数：每个输出在全部路径（含提前返回）上赋值。
 * 错误码    : 16#0001_03C1 填充字符为空（已按空格降级）——信息级
 *             16#0001_03C2 保留禁用（不得挪用，本件零赋值）
 * 码位总账  : 16#0001_03C1 用 ｜ 16#0001_03C2 预留
 * 修改记录  : v1.0.0 R26 初版
 *==============================================================================*)
FUNCTION FC_DL_StringPad : BOOL
VAR_INPUT
    sIn         : STRING; // 源字符串 / Source string
    sPadChar    : STRING; // 填充字符（取首字符，空则降级空格）/ Pad char (first char, empty degrades to space)
    nTargetLen  : UINT;   // 目标长度 0~255 / Target length 0 to 255
    eSide       : E_DL_PadSide; // 填充侧别：左/右/居中 / Pad side: left, right or center
END_VAR
VAR_OUTPUT
    sOut        : STRING; // 填充结果字符串 / Padded result string
    bTruncated  : BOOL;  // 发生截断（源超长或目标超界钳 255）/ Truncation occurred
    eErr        : UDINT;  // 本周期错误码，0=无错 / Error code this cycle, 0 = none
END_VAR
VAR
    iTarget : INT; // 目标长度有效值（钳 255 后）/ Effective target length after clamp
    iSrcLen : INT; // 源串实际长度 / Actual source length
    iLeft   : INT; // 左侧填充字符数 / Left pad char count
    iRight  : INT; // 右侧填充字符数 / Right pad char count
    i       : INT; // 循环游标 / Loop cursor
    sPadOne : STRING; // 单个填充字符（首字符或降级空格）/ Single pad char
    sPadL   : STRING; // 左侧填充串 / Left pad string
    sPadR   : STRING; // 右侧填充串 / Right pad string
END_VAR

// ---------- 全路径赋值原则：先给输出安全缺省 ----------
sOut       := '';
bTruncated := FALSE;
eErr       := 0;
FC_DL_StringPad := TRUE; // 函数返回值：TRUE=已执行（防御缺省）/ Function result: TRUE = executed

// ---------- 目标长度钳位：超 255 显式截断标记 ----------
IF nTargetLen > 255 THEN
    iTarget    := 255;                        // 超界钳 255 / Clamp over-range to 255
    bTruncated := TRUE;                       // 显式置截断标志，禁静默回夹 / Explicit truncation flag
ELSE
    iTarget := UINT_TO_INT(nTargetLen);       // 合法目标长度 / Legal target length
END_IF

// ---------- 填充字符取首字符；空串降级为空格并置信息码 ----------
IF LEN(sPadChar) <= 0 THEN
    sPadOne := ' ';                           // 降级为空格 / Degrade to space
    eErr    := 16#0001_03C1;                  // 信息级：填充字符为空已降级 / info: empty pad char degraded
ELSE
    sPadOne := MID(sPadChar, 1, 1);           // 取首字符 / Take first char
END_IF

// ---------- 源串长度与超长截断 ----------
iSrcLen := LEN(sIn);
IF iSrcLen > iTarget THEN
    sOut       := LEFT(sIn, iTarget);         // 按目标长度截断 / Truncate to target
    bTruncated := TRUE;                       // 显式截断标志 / Explicit truncation flag
    RETURN;                                   // 提前返回路径：输出已全赋值 / Early return: outputs all assigned
END_IF

// ---------- 按侧别计算左右填充量 ----------
CASE eSide OF
    E_DL_PadSide.eLeft:                       // 左填充 / Left padding
        iLeft  := iTarget - iSrcLen;          // 全部填左侧 / All padding on the left
        iRight := 0;
    E_DL_PadSide.eRight:                      // 右填充 / Right padding
        iLeft  := 0;
        iRight := iTarget - iSrcLen;          // 全部填右侧 / All padding on the right
    E_DL_PadSide.eCenter:                     // 居中：奇偶差一填左侧 / Center: odd remainder goes left
        iLeft  := (iTarget - iSrcLen + 1) / 2; // 左侧含奇余 / Left side takes odd remainder
        iRight := (iTarget - iSrcLen) / 2;     // 右侧取偶商 / Right side takes even quotient
    ELSE                                      // 非法侧别防御降级为右填充 / Illegal side degrades to right
        iLeft  := 0;
        iRight := iTarget - iSrcLen;
END_CASE

// ---------- 逐字符构造填充串（标准 CONCAT，避免方言拼接符） ----------
sPadL := '';
FOR i := 1 TO iLeft DO
    sPadL := CONCAT(sPadL, sPadOne);          // 累积左侧填充 / Accumulate left padding
END_FOR
sPadR := '';
FOR i := 1 TO iRight DO
    sPadR := CONCAT(sPadR, sPadOne);          // 累积右侧填充 / Accumulate right padding
END_FOR

// ---------- 组装输出：左填充串 + 源串 + 右填充串 ----------
IF iLeft > 0 THEN
    sOut := CONCAT(sPadL, sIn);               // 先贴左填充 / Attach left padding first
ELSE
    sOut := sIn;                              // 无左填充直接用源串 / No left pad, use source
END_IF
IF iRight > 0 THEN
    sOut := CONCAT(sOut, sPadR);              // 再贴右填充 / Then attach right padding
END_IF

END_FUNCTION

(* ---- FC_DL_StringReplaceAll.st ---- *)
(*==============================================================================
 * 组件名称 (Component)  : FC_DL_StringReplaceAll
 * 所属子库 (Sublibrary) : DL_MathData
 * 当前版本 (Version)    : 1.0.1
 * 兼容性   (Platform)   : CODESYS 3.5 / TwinCAT 3 / 汇川 InoProShop / Machine Expert
 *                         仅依赖 Standard.library 标准串函数（LEN / FIND / LEFT / MID / CONCAT）
 * 功能描述 (Function)   : 定长字符串内「全部出现」的子串替换，一次调用给出替换次数、
 *                         结果串与截断标志。用于条码前缀规范化、报表模板占位符替换
 *                         （百分号包裹的批次号与日期占位符）、设备商旧机型代号批量改新代号。
 *                         现场手写 WHILE + FIND + DELETE + INSERT 的典型事故是「替换串里
 *                         含模式串」时缓冲自增长、永不退出扫描，本件用「替换后游标跳到
 *                         插入段之后」的推进律从算法层消灭该类死循环，并叠加次数上限与
 *                         守卫计数器两道闸。
 * 出口契约 (Exit)       : 函数返回值 = 实际替换次数（与出口 nReplaced 同值）；异常路径返回 0。
 *                         任何路径（含早退）sResult 均有确定内容，绝不返回未初始化串。
 * 开源溯源 (Origin)     : 来源标签 lgf-datahandling。许可证：LGF 为免费闭源发布，未取得源码，
 *                         不构成衍生作品。借鉴点仅为「Data Handling 组把 FIFO/LIFO、数组检索、
 *                         排序、字符串并列成数据操作族」的分类骨架，以及字符串族「定长缓冲 +
 *                         原地操作、不做动态分配」的参数域约定。
 *                         clean-room 独立实现：算法、切分策略、游标推进律、计数语义、错误码
 *                         全部自有，零代码行、零注释、零结构体复制。
 * 码位说明 (Codes)      : 信息级 16#0001_0130（模式串为空）/ 0131（达替换次数上限）/
 *                         0132（结果被长度上限截断）/ 0133（长度参数越界已钳位）。
 *                         共 4 码，全部落在 R12 计划第 1.2 节分配给本件的码段内，无段外码。
 * 依赖     (Depends)    : 无 DL_ 内部依赖；Standard.library: LEN / FIND / LEFT / MID / CONCAT
 * 红线自检 (Redline)    : 1 ✓ 零全局变量表依赖、零外部变量声明、零物理地址
 *                         2 ✓ 纯 IEC 61131-3 跨平台语法，无指针、无厂商库
 *                         3 ✓ 模式空硬闸、数组与串长先判界、每轮回夹、双闸防死循环
 *                         4 ✓ 全变量中英双语同行注释
 *                         5 N/A 纯函数无状态机 ｜ 6 N/A 无定时器与边沿实例
 *                         7 ✓ END_FUNCTION 位于文件最后有效行
 * 规格偏离留档 (Deviation):
 *   D1 计划 3.6 节把 bValid 定义为「模式串非空且长度参数合法」。本实现多收一环：
 *      达替换次数上限（码 0131，结果不完整）时 bValid 亦为假。理由：bValid 在本库
 *      统一承载「结果可否直接采信」，不完整的替换结果采信即等于静默丢字段；
 *      完整性细粒度判据由调用方读 uErrorId 与 bTruncated 取得。
 * 修订历史 (Revision)   :
 *   2026-11-15  v1.0.0  首版入库（R12 · Level 0 DL_MathData 字符串族）
 *   2026-11-15  v1.0.1  终审定点修复 A-D01：拼接长度超串型上限（255）时原实现由
 *      LEFT 静默回夹，bTruncated 与 0132 永不置位（验收向量 V5 期望的截断标志恒假）；
 *      补「拼接长度预判」，超限即置 bTruncated 与 0132，杜绝静默丢字符
 *============================================================================*)
FUNCTION FC_DL_StringReplaceAll : INT
VAR_INPUT
    sSource      : STRING(255);          // 源串，最长 255 字符 / Source string, up to 255 characters
    sPattern     : STRING(32);           // 被替换子串，长度 0 视为非法 / Pattern to replace, empty is illegal
    sReplace     : STRING(64);           // 替换子串，允许为空（即删除） / Replacement, empty means delete
    nMaxReplace  : INT := 32;            // 替换次数上限 [次]，域 0~255，0 = 不限 / Replacement limit, zero means unlimited
    nMaxLen      : INT := 255;           // 结果串长度上限 [字符]，域 1~255 / Result length limit, 1..255
END_VAR
VAR_OUTPUT
    sResult      : STRING(255);          // 替换结果，超长时按 nMaxLen 截断 / Result, truncated to nMaxLen
    nReplaced    : INT;                  // 实际替换次数 [次] / Replacement count
    bTruncated   : BOOL;                 // 结果被长度上限截断 TRUE / Result was truncated
    uErrorId     : UDINT;                // 事件码，0 = 无事件 / Event code, zero means none
    bValid       : BOOL;                 // 模式串非空、长度参数未钳位且未达替换次数上限 = TRUE（结果可直接采信） / Pattern non-empty, lengths legal and the count limit not hit, the result may be trusted as is
END_VAR
VAR
    sBuf         : STRING(255);          // 工作缓冲，逐轮就地改写 / Working buffer, rewritten in place
    sHead         : STRING(255);         // 本次替换位置之前的头部片段 / Head fragment before the hit
    sTail        : STRING(255);          // 本次替换位置之后的尾部片段 / Tail fragment after the hit
    sScan        : STRING(255);          // 查找窗口，从 nSearchFrom 起的剩余串 / Search window starting at nSearchFrom
    nPos         : INT;                  // 当前命中位置，1 起，0 = 未命中 [字符位] / Current hit position, one based
    nSearchFrom  : INT;                  // 下一轮查找起点，1 起 [字符位] / Next search start position
    nLenBuf      : INT;                  // 当前缓冲长度 [字符] / Current buffer length
    nLenPat      : INT;                  // 模式串长度 [字符] / Pattern length
    nLenRep      : INT;                  // 替换串长度 [字符] / Replacement length
    nTailStart   : INT;                  // 尾部片段起始位置 [字符位] / Tail fragment start position
    nMaxRepUse   : INT;                  // 生效替换次数上限 [次] / Effective replacement limit
    nMaxLenUse   : INT;                  // 生效结果长度上限 [字符] / Effective result length limit
    nGuard       : DINT;                 // 循环守卫，防串函数异常导致死循环 / Loop guard against endless looping
END_VAR
VAR CONSTANT
    DL_STR_MAX   : INT  := 255;          // 单字节串长度上限，与类型声明一致 [字符] / Single byte string ceiling
    DL_PAT_MAX   : INT  := 32;           // 模式串长度上限，与入参声明一致 [字符] / Pattern ceiling
    DL_REP_MAX   : INT  := 64;           // 替换串长度上限，与入参声明一致 [字符] / Replacement ceiling
    DL_GUARD_MAX : DINT := 512;          // 循环守卫上限 [次] / Loop guard limit
END_VAR

(*------------------------------------------------------------------------------
 * 段 1｜结果预置（P-01 范式）：先给全部出口与全部中间量确定值
 *      Safe preset: every output and every intermediate gets a defined value
 *-----------------------------------------------------------------------------*)
FC_DL_StringReplaceAll := 0;
sResult    := '';
nReplaced  := 0;
bTruncated := FALSE;
uErrorId   := 16#0000_0000;
bValid     := FALSE;
sBuf       := '';
sHead      := '';
sTail      := '';
sScan      := '';
nPos       := 0;
nSearchFrom := 1;
nLenBuf    := 0;
nLenPat    := 0;
nLenRep    := 0;
nTailStart := 0;
nMaxRepUse := 0;
nMaxLenUse := 1;
nGuard     := 0;

(*------------------------------------------------------------------------------
 * 段 2｜参数闸门：串长快照 + 两个长度上限钳位（信息级，钳位后照常执行）
 *      Parameter gates: string snapshots and the two length clamps (informational)
 *-----------------------------------------------------------------------------*)
nLenPat := LEN(sPattern);
IF nLenPat > DL_PAT_MAX THEN
    nLenPat := DL_PAT_MAX;
END_IF
nLenRep := LEN(sReplace);
IF nLenRep > DL_REP_MAX THEN
    nLenRep := DL_REP_MAX;
END_IF

nMaxRepUse := nMaxReplace;
IF nMaxRepUse < 0 THEN
    nMaxRepUse := 0;
    uErrorId := 16#0001_0133;
ELSIF nMaxRepUse > DL_STR_MAX THEN
    nMaxRepUse := DL_STR_MAX;
    IF uErrorId = 16#0000_0000 THEN
        uErrorId := 16#0001_0133;
    END_IF
END_IF
IF nMaxRepUse = 0 THEN
    nMaxRepUse := DL_STR_MAX;
END_IF

nMaxLenUse := nMaxLen;
IF nMaxLenUse < 1 THEN
    nMaxLenUse := 1;
    IF uErrorId = 16#0000_0000 THEN
        uErrorId := 16#0001_0133;
    END_IF
ELSIF nMaxLenUse > DL_STR_MAX THEN
    nMaxLenUse := DL_STR_MAX;
    IF uErrorId = 16#0000_0000 THEN
        uErrorId := 16#0001_0133;
    END_IF
END_IF

bValid := (uErrorId = 16#0000_0000);
sBuf   := LEFT(sSource, DL_STR_MAX);

(*------------------------------------------------------------------------------
 * 段 3｜模式串硬闸：长度 0 直接早退，绝不进入查找循环
 *      Hard gate on the pattern: a zero length pattern never reaches the loop
 *      空模式在 FIND 上的行为跨平台不一致，且会让游标推进律失效，必须在算法入口拦死
 *      An empty pattern makes FIND platform dependent and breaks cursor advance
 *-----------------------------------------------------------------------------*)
IF nLenPat <= 0 THEN
    bValid   := FALSE;
    uErrorId := 16#0001_0130;
ELSE

    (*--------------------------------------------------------------------------
     * 段 4｜主替换循环：三闸并行 —— 次数上限、守卫计数、游标只前进
     *      Main replace loop guarded by the count limit, the guard counter and a
     *      strictly advancing cursor
     *      切分口径：头部保留 + 替换串 + 尾部保留，拼装后立即按串上限回夹
     *      Split policy: head kept, replacement inserted, tail kept, then re-clamped
     *      回夹前必须预判长度：静默回夹等于丢字符，bTruncated 与 0132 必须同时置位
     *      The length is predicted before clamping so truncation is never silent
     *-----------------------------------------------------------------------*)
    nSearchFrom := 1;
    nReplaced   := 0;
    nGuard      := 0;

    WHILE (nReplaced < nMaxRepUse) AND (nGuard < DL_GUARD_MAX) DO
        nGuard  := nGuard + 1;
        nLenBuf := LEN(sBuf);
        nPos    := 0;

        IF (nSearchFrom >= 1) AND (nSearchFrom <= nLenBuf) THEN
            sScan := MID(sBuf, nLenBuf - nSearchFrom + 1, nSearchFrom);
            nPos  := FIND(sScan, sPattern);
            IF nPos > 0 THEN
                nPos := nPos + nSearchFrom - 1;
            END_IF
        END_IF

        IF nPos <= 0 THEN
            EXIT;
        END_IF

        IF nPos > 1 THEN
            sHead := LEFT(sBuf, nPos - 1);
        ELSE
            sHead := '';
        END_IF

        nTailStart := nPos + nLenPat;
        IF nTailStart <= nLenBuf THEN
            sTail := MID(sBuf, nLenBuf - nTailStart + 1, nTailStart);
        ELSE
            sTail := '';
        END_IF

        (* 拼接长度预判：超出串型上限即属截断，先置标志与事件码，绝不静默丢字符 *)
        (* Predict the joined length: exceeding the string ceiling is a truncation *)
        IF (LEN(sHead) + nLenRep + LEN(sTail)) > DL_STR_MAX THEN
            bTruncated := TRUE;
            IF uErrorId = 16#0000_0000 THEN
                uErrorId := 16#0001_0132;
            END_IF
        END_IF
        sBuf := CONCAT(sHead, sReplace);
        sBuf := CONCAT(sBuf, sTail);
        sBuf := LEFT(sBuf, DL_STR_MAX);

        nReplaced := nReplaced + 1;

        (* 游标跳到「已插入替换串之后」：替换串含模式串时天然跳过新插入段 *)
        (* Cursor jumps past the inserted replacement: self growing patterns are safe *)
        nSearchFrom := nPos + nLenRep;
        IF nSearchFrom < 1 THEN
            nSearchFrom := 1;
        END_IF
    END_WHILE;

    (*--------------------------------------------------------------------------
     * 段 5｜上限判定：达到次数上限且剩余串内仍有模式串，说明结果不完整
     *      Limit verdict: hitting the count limit with the pattern still present
     *      means the result is incomplete and must be reported, never silently cut
     *-----------------------------------------------------------------------*)
    nLenBuf := LEN(sBuf);
    IF nReplaced >= nMaxRepUse THEN
        nPos := 0;
        IF (nSearchFrom >= 1) AND (nSearchFrom <= nLenBuf) THEN
            sScan := MID(sBuf, nLenBuf - nSearchFrom + 1, nSearchFrom);
            nPos  := FIND(sScan, sPattern);
        END_IF
        IF nPos > 0 THEN
            bValid := FALSE;
            IF uErrorId = 16#0000_0000 THEN
                uErrorId := 16#0001_0131;
            END_IF
        END_IF
    END_IF

END_IF

(*------------------------------------------------------------------------------
 * 段 6｜结果截断（两条路径共用）：超长按上限裁剪并置标志，事件码首事件优先
 *      Shared truncation step: crop to the limit and keep the first event code
 *-----------------------------------------------------------------------------*)
nLenBuf := LEN(sBuf);
IF nLenBuf > nMaxLenUse THEN
    sBuf       := LEFT(sBuf, nMaxLenUse);
    bTruncated := TRUE;
    IF uErrorId = 16#0000_0000 THEN
        uErrorId := 16#0001_0132;
    END_IF
END_IF

(*------------------------------------------------------------------------------
 * 段 7｜结果落地：返回值与出口同源，保证「同入参同结果」的可重入语义
 *      Result publication: the return value and the output share one source
 *-----------------------------------------------------------------------------*)
sResult := sBuf;
FC_DL_StringReplaceAll := nReplaced;
END_FUNCTION
